(* IEC 61131-3 sources: daoli-st-library/DL_Algo (part 13) *)

(* ---- FB_DL_FirFilter.st ---- *)
(*==============================================================================
 * 组件名称 (Component)  : FB_DL_FirFilter
 * 所属子库 (Sublibrary) : DL_Algo
 * 当前版本 (Version)    : 1.0.0
 * 兼容性   (Platform)   : CODESYS 3.5+ / TwinCAT 3 / 汇川 InoProShop / 施耐德 Machine Expert
 *                         仅依赖 Standard.library（ABS），零厂商私有库
 * 功能描述 (Function)   : N 阶 FIR 直接型滤波器：抽头系数 aCoeffs[0..nTaps−1]
 *                         （aCoeffs[0] 对应最新样本，倒序卷积）：
 *                           fFiltered = Σ aCoeffs[k] × aHist[k]，k ∈ [0, nTaps−1]
 *                         样本入栈做循环移位（自深至浅倒序拷贝，防越界覆盖）。
 *                         系数和归一校验：|ΣaCoeffs − 1| < 1E-6，破约 → 锁存
 *                         故障 eCoeffSum（直流增益 ≠ 1 会引入稳态偏差，锁存
 *                         冻结输出）；N 阶钳位 [1,16]，越界钳位并置信息码
 *                         eTapsClamp；非有限样本跳过入栈并置信息码 eSampleSkip。
 * 接口     (Interface)  : 输入 fSample 输入样本、aCoeffs 抽头系数表（定长
 *                         0..15）、nTaps 有效抽头数（钳位 1~16）、bReset 复位；
 *                         输出 fFiltered 滤波输出、fCoeffSum 实测系数和
 *                         （诊断透读）、eErrCode 错误码、bError 故障标志。
 * 边界     (Boundary)   : ① **属主边界（写死）：本件只做 FIR 直接型卷积，不做
 *                         系数设计、不做 IIR 递推**；系数设计离线完成。
 *                         ② 移位：FOR 自深至浅倒序拷贝 aHist[i] := aHist[i−1]
 *                         （i ∈ [1, nTaps−1]，界宽 = 钳位后 nTaps，无越界），
 *                         aHist[0] := fSample 唯一写入点。
 *                         ③ 卷积求和界宽 = 钳位后 nTaps；aHist 尾部旧样本
 *                         （从未填充）为初值 0，首窗输出为尾零卷积（头注释
 *                         声明：上电启动期输出按零历史卷积，非异常）。
 *                         ④ 系数和归一校验在每次 nTaps 钳位后按活动抽头重算；
 *                         破约锁存后冻结输出 0（安全侧），解除沿 = bReset
 *                         上升沿（故障级码配对 bError，R45）。
 *                         ⑤ 非有限判据（R79 双判）：样本跳过（不入栈不卷积），
 *                         系数域闸含逐系数非有限判（系数 NaN 直接判归一破约
 *                         路径覆盖，另设显式非有限分支置 eCoeffSum）。
 *                         ⑥ 零全局耦合（无 GVL / VAR_EXTERNAL / 物理地址）。
 * 分工声明 (Scope)      : 与 `FB_DL_MovingAverage` 分工：等权滑动平均（FIR 特例）
 *                         归那件、任意系数 FIR 归本件；与 `FB_DL_LowPassFilter`
 *                         分工：IIR 单极点归那件。
 * 来源标签 (Source Tag) : 自研线（FIR 直接型为公开 DSP 结构 clean-room）
 * 码表     (Codes)      : 本件不占用任何全局数字码位。出口为 LREAL 组 +
 *                         ENUM 错误码；数字码位待主控收口阶段统一派号。
 * 红线自检 (Redline)    : R1 ✓ 零 GVL/VAR_EXTERNAL ｜ R2 ✓ 零 %I/%Q/%M ｜ R3 ✓ 纯 IEC 61131-3
 *                         R4 ✓ 移位界宽钳位 + 归一校验锁存 + 非有限跳过 ｜ R5 ✓ 声明逐行同行双语注释
 *                         R6 N/A（无 ENUM 状态机） ｜ R7 ✓ 一 R_TRIG 段 0 无条件刷新
 * 修订历史 (Revision)   : 2026-11-20  v1.0.0  R50 首版（批次 2 · 序号 9）
 * 验收向量 (Acceptance) : ① nTaps=2，aCoeffs=[0.5, 0.5]（Σ=1.0 过闸）：样本
 *                         序列 10, 20 → 首拍输出 0.5×10+0.5×0 = 5.0（零历史），
 *                         次拍 0.5×20+0.5×10 = 15.0，eOk；② nTaps=20 → 钳位
 *                         16，eTapsClamp；③ aCoeffs=[0.6, 0.5]（Σ=1.1）→
 *                         |1.1−1|=0.1 ≥ 1E-6 → 锁存 eCoeffSum，输出 0；
 *                         ④ 样本 NaN → uSkip 不入栈，eSampleSkip，输出不变。
 *==============================================================================*)

(*-----------------------------------------------------------------------------
 * 枚举: E_DL_FirErr（错误码；信息级不置 bError，故障级恒伴 bError=TRUE）
 *----------------------------------------------------------------------------*)
TYPE E_DL_FirErr :
(
    eOk          := 0,   // 正常 / Normal
    eCoeffSum    := 1,   // 故障级：系数和归一破约（|Σ−1| ≥ 1E-6 或含非有限） / Fault: coefficient sum not unity
    eTapsClamp   := 2,   // 信息级：抽头数越界已钳位 [1,16] / Info: tap count clamped
    eSampleSkip  := 3    // 信息级：样本非有限已跳过 / Info: non-finite sample skipped
);
END_TYPE

FUNCTION_BLOCK FB_DL_FirFilter
VAR_INPUT
    fSample : LREAL := 0.0;                    // 输入样本 [工程单位] / Input sample
    aCoeffs : ARRAY[0..15] OF LREAL;           // 抽头系数表（[0] 对应最新样本） [-] / Tap coefficients, newest-first
    nTaps   : UDINT := 4;                      // 有效抽头数，域 [1,16]（越界钳位） [个] / Active tap count
    bReset  : BOOL := FALSE;                   // 复位，上升沿清组态锁存与历史栈 [-] / Reset, rising edge clears latch and history
END_VAR
VAR_OUTPUT
    fFiltered  : LREAL;                        // 滤波输出 [工程单位] / Filtered output
    fCoeffSum  : LREAL;                        // 实测活动抽头系数和（诊断透读） [-] / Measured coefficient sum
    eErrCode   : E_DL_FirErr;                  // 错误码出口 / Error code outlet
    bError     : BOOL;                         // 故障标志（归一破约锁存） [-] / Error flag, latched
END_VAR
VAR
    _aHist    : ARRAY[0..15] OF LREAL;         // 历史样本栈（aHist[0] 最新，初值零历史） / History stack, newest first
    _nTaps    : DINT;                          // 钳位后抽头数 [个] / Clamped tap count
    _fSum     : LREAL;                         // 系数和累计中间量 [-] / Coefficient sum intermediate
    _fAcc     : LREAL;                         // 卷积累计中间量 [工程单位] / Convolution accumulator
    _bClamp   : BOOL;                          // 本拍发生抽头钳位 [-] / Tap clamp this scan
    _bNonFin  : BOOL;                          // 样本非有限当拍量 [-] / Sample non-finite this scan
    _bCoefBad : BOOL;                          // 系数归一破约当拍量 [-] / Coefficient sum violation this scan
    _bErrLatch: BOOL;                          // 归一破约锁存位（解除沿 = bReset 上升沿） / Latched coeff-sum fault
    i         : DINT;                          // 移位/卷积循环索引 / Shift and convolution loop index
    rtReset   : R_TRIG;                        // 复位沿实例，段 0 无条件调用 / Reset edge instance
END_VAR
VAR CONSTANT
    DL_FIR_NMAX   : DINT  := 16;               // 抽头定长上限 [个] / Tap count ceiling
    DL_FIR_NMIN   : DINT  := 1;                // 抽头数下限 [个] / Tap count floor
    DL_FIR_SUMTOL : LREAL := 1.0E-6;           // 系数和归一容差 [-] / Coefficient sum tolerance
    DL_FIR_ONE    : LREAL := 1.0;              // 归一目标值 [-] / Unity target
    DL_FIR_ZERO   : LREAL := 0.0;              // 判零与安全侧基准 / Zero base and safe value
END_VAR

(* —— 段 0：抽头钳位 + 非有限判 + 沿刷新 —— *)
_bClamp := FALSE;                              // 钳位量预清 / Clamp preset
_nTaps := UDINT_TO_DINT(nTaps);                // 抽头数转 DINT（越界由下步钳位） / Convert tap count
IF _nTaps > DL_FIR_NMAX THEN
    _nTaps := DL_FIR_NMAX;                     // 上越界钳 16 / Clamp high
    _bClamp := TRUE;                           // 记钳位 / Mark clamp
END_IF
IF _nTaps < DL_FIR_NMIN THEN
    _nTaps := DL_FIR_NMIN;                     // 下越界钳 1 / Clamp low
    _bClamp := TRUE;                           // 记钳位 / Mark clamp
END_IF
_bNonFin := (fSample <> fSample) OR ((fSample - fSample) <> DL_FIR_ZERO);   // 样本非有限（R79 双判） / Sample non-finite
rtReset(CLK := bReset);                        // 复位沿，每拍必调 / Reset edge, every scan

(* —— 段 1：复位沿（清锁存与历史栈） —— *)
IF rtReset.Q THEN
    _bErrLatch := FALSE;                       // 清归一破约锁存（R188 声明：解除沿 = bReset 上升沿） / Clear latch
    FOR i := 0 TO (DL_FIR_NMAX - 1) DO
        _aHist[i] := DL_FIR_ZERO;              // 清历史栈（零历史重启） / Clear history stack
    END_FOR
END_IF

(* —— 段 2：系数和归一校验（按钳位后活动抽头重算；含系数非有限判） —— *)
_fSum := DL_FIR_ZERO;                          // 系数和起步 0 / Sum start zero
FOR i := 0 TO (_nTaps - 1) DO
    _fSum := _fSum + aCoeffs[i];               // 活动抽头逐项累计 / Sum active taps
END_FOR
fCoeffSum := _fSum;                            // 透读出口 / Readout outlet
IF (_fSum <> _fSum) OR ((_fSum - _fSum) <> DL_FIR_ZERO)
   OR (ABS(_fSum - DL_FIR_ONE) >= DL_FIR_SUMTOL) THEN
    _bCoefBad := TRUE;                         // 归一破约（含系数 NaN 令和失效） / Sum violation
ELSE
    _bCoefBad := FALSE;                        // 过闸 / Pass
END_IF
IF _bCoefBad AND (NOT _bErrLatch) THEN
    _bErrLatch := TRUE;                        // 锁存（R188） / Latch
END_IF

(* —— 段 3：样本入栈（循环移位倒序拷贝，防越界；故障期/非有限期不入栈） —— *)
IF (NOT _bErrLatch) AND (NOT _bNonFin) THEN
    FOR i := (_nTaps - 1) TO DL_FIR_NMIN BY -1 DO
        _aHist[i] := _aHist[i - 1];            // 倒序拷贝（自深至浅，界宽=nTaps） / Shift down, newest-first
    END_FOR
    _aHist[0] := fSample;                      // 最新样本入栈（唯一写入点） / Push newest sample
END_IF

(* —— 段 4：卷积输出（故障安全侧 0；正常域按活动抽头求和） —— *)
IF _bErrLatch THEN
    fFiltered := DL_FIR_ZERO;                  // 归一破约冻结输出 0（安全侧，头注释④） / Frozen zero output
ELSE
    _fAcc := DL_FIR_ZERO;                      // 卷积累计起步 0 / Accumulator start
    FOR i := 0 TO (_nTaps - 1) DO
        _fAcc := _fAcc + aCoeffs[i] * _aHist[i];   // 倒序卷积逐项 / Tap-wise convolution
    END_FOR
    fFiltered := _fAcc;                        // 滤波输出 / Filtered outlet
END_IF

(* —— 段 5：出口单点映射（错误码归约，R191） —— *)
IF _bErrLatch THEN
    bError := TRUE;                            // 故障标志（R45 配对） / Error flag
    eErrCode := E_DL_FirErr.eCoeffSum;         // 故障级码 / Fault code
ELSE
    bError := FALSE;                           // 无故障级条件 / No fault
    IF _bNonFin THEN
        eErrCode := E_DL_FirErr.eSampleSkip;   // 信息级：样本跳过 / Info: skipped
    ELSIF _bClamp THEN
        eErrCode := E_DL_FirErr.eTapsClamp;    // 信息级：抽头钳位 / Info: clamped
    ELSE
        eErrCode := E_DL_FirErr.eOk;           // 正常 / Normal
    END_IF
END_IF

END_FUNCTION_BLOCK

(* ---- FB_DL_FirstOrderIdent.st ---- *)
(*
  Name        : FB_DL_FirstOrderIdent
  Category    : DL_Algo
  Version     : 1.0.0
  Purpose     : 一阶加纯滞后（FOPDT）阶跃响应回归：阶跃前后双特征点三点法估增益/时间常数/纯滞后，供自整定与 Smith 补偿取参；/ FOPDT step-response regression: two feature points before and after the step estimate gain, time constant and dead time for auto-tuning and Smith predictor
  溯源        : 自研（与 PRBS/继电器整定/扫频激励源配套），clean-room 实现
  Boundary    : ① 阶跃幅值/采样周期/窗长三重域闸，任一越域锁存故障；
                ② 辨识窗须含阶跃前稳态（>= 8 有效拍均值）与阶跃后 28.3%/63.2% 两特征点，缺任一 → 有效性 FALSE 不出参数（信息级）；
                ③ 三点法公式全代数无迭代（增益分母 = 阶跃幅值，已过正域闸；除子常量均非零）；
                ④ 非有限测量该拍不入辨识窗（窗计数暂停非快进，防污染统计）；
                ⑤ 输出 K/T/θ 非负域钳位，θ 上限 = 辨识窗时长（防无滞后误设大滞后）；
                ⑥ 本件为辨识观测层，不输出任何控制量（属主边界）。
*)
TYPE E_DL_FoiState :
(
    eIdle  := 0,                             (* 未辨识 / Not identifying *)
    eWait  := 10,                            (* 阶跃前稳态采集 / Pre-step steady sampling *)
    ePost  := 20,                            (* 阶跃后窗采集 / Post-step window sampling *)
    eReady := 30,                            (* 辨识完成（有效性查 bValid） / Finished, see bValid *)
    eFault := 90                             (* 故障锁存相 / Fault latched *)
);
END_TYPE

TYPE E_DL_FoiCause :
(
    eNone      := 0,                         (* 无成因 / No cause *)
    eCfgIllegal:= 1,                        (* 组态非法：幅值/周期/窗长越域 / Illegal config *)
    eNoFeat    := 2,                        (* 信息级：缺稳态/特征点或增益反号 / Info: feature missing *)
    ePhaseBad  := 3                         (* 非法相位兜底 / Illegal phase fallback *)
);
END_TYPE

FUNCTION_BLOCK FB_DL_FirstOrderIdent
VAR_INPUT
    fMeas   : REAL := 0.0;                   (* 回路测量值（任意工程量）[-] / Loop measurement *)
    fStepAmp: REAL := 10.0;                  (* 阶跃幅值，域 > 0 [工程单位] / Step amplitude *)
    tSample : TIME := T#100MS;               (* 采样周期，域 > T#0S [ms] / Sampling period *)
    nWin    : INT := 128;                    (* 阶跃后窗长，域 20..256 [拍] / Post-step window length *)
    bStart  : BOOL := FALSE;                 (* 启动辨识命令，上升沿进入稳态采集 [-] / Start command *)
    bEnable : BOOL := TRUE;                  (* 使能 [-] / Enable *)
    bReset  : BOOL := FALSE;                 (* 复位命令，上升沿清故障与结果 [-] / Reset command *)
END_VAR
VAR_OUTPUT
    fK      : REAL;                          (* 增益出口 = 稳态增量 / 阶跃幅值 [-] / Gain outlet *)
    fTau    : REAL;                          (* 时间常数出口 [s] / Time constant outlet *)
    fTheta  : REAL;                          (* 纯滞后出口（非负，上限 = 窗时长）[s] / Dead time outlet *)
    bValid  : BOOL;                          (* 结果有效性出口 [-] / Result validity *)
    nSamples: INT;                           (* 阶跃后窗内有效样本数 [拍] / Valid samples in window *)
    eState  : E_DL_FoiState;                 (* 状态出口 / State outlet *)
    eCause  : E_DL_FoiCause;                 (* 成因出口（R190 归因唯一） / Cause outlet *)
    bError  : BOOL;                          (* 故障锁存标志 [-] / Fault latch flag *)
END_VAR
VAR
    _eState : E_DL_FoiState := E_DL_FoiState.eIdle;  (* 内部相位（CASE 唯一写入目标） / Internal phase *)
    _eCause : E_DL_FoiCause := E_DL_FoiCause.eNone;  (* 成因锁存量 / Latched cause *)
    rtStart : R_TRIG;                        (* 启动沿实例，段 0 无条件调用 / Start edge instance *)
    rtReset : R_TRIG;                        (* 复位沿实例，段 0 无条件调用 / Reset edge instance *)
    _bFault : BOOL;                          (* 故障锁存位 / Latched fault bit *)
    _bCfgBad: BOOL;                          (* 组态非法当拍量 / Illegal config this scan *)
    _bFin   : BOOL;                          (* 测量有限性当拍量（边界④） / Measurement finiteness *)
    _nWinE  : INT;                           (* 钳位后生效窗长 [拍] / Effective window length *)
    _nPreN  : INT;                           (* 稳态已采有效拍数 [拍] / Pre samples collected *)
    _fPreSum: REAL;                          (* 稳态样本累加和 [工程单位] / Pre samples sum *)
    _fY0    : REAL;                          (* 阶跃前稳态均值 [工程单位] / Baseline mean *)
    _nRecN  : INT;                           (* 窗内已收有效样本数 [拍] / Window samples count *)
    _aRec   : ARRAY[1..256] OF REAL;         (* 窗内样本记录（连续有效区）[工程单位] / Window sample record *)
    _fYinf  : REAL;                          (* 窗末稳态均值 [工程单位] / Final steady mean *)
    _fDelta : REAL;                          (* 稳态增量中间量 [工程单位] / Steady delta *)
    _fKI    : REAL;                          (* 增益中间量 [-] / Gain intermediate *)
    _fT1    : REAL;                          (* 28.3% 特征时刻 [s] / Feature time 1 *)
    _fT2    : REAL;                          (* 63.2% 特征时刻 [s] / Feature time 2 *)
    _fTauI  : REAL;                          (* 时间常数中间量 [s] / Tau intermediate *)
    _fThI   : REAL;                          (* 滞后中间量 [s] / Theta intermediate *)
    _i      : INT;                           (* 窗扫描游标 [拍] / Window scan cursor *)
    _fDtSec : REAL;                          (* 采样周期秒值，域 > eps [s] / Sampling period seconds *)
END_VAR
VAR CONSTANT
    DL_FOI_NPRE   : INT  := 8;               (* 阶跃前稳态最少有效拍数（边界②）[拍] / Pre-step minimum samples *)
    DL_FOI_NTAIL  : INT  := 8;               (* 窗末稳态平均样本数 [拍] / Tail averaging samples *)
    DL_FOI_WMIN   : INT  := 20;              (* 窗长下限（边界①）[拍] / Window lower bound *)
    DL_FOI_WMAX   : INT  := 256;             (* 窗长上限（数组容量）[拍] / Window upper bound *)
    DL_FOI_EPS    : REAL := 1.0E-6;          (* 判零容差 [-] / Epsilon *)
    DL_FOI_L1     : REAL := 0.283;           (* 特征点 1 归一化水平（1-exp(-1/3)）[-] / Feature level 1 *)
    DL_FOI_L2     : REAL := 0.632;           (* 特征点 2 归一化水平（1-exp(-1)）[-] / Feature level 2 *)
    DL_FOI_STEPDET: REAL := 0.1;             (* 阶跃检测阈（幅值占比）[-] / Step detect threshold *)
END_VAR

(* —— 段 0：当拍判据派生 + 实例无条件刷新（R228A） —— *)
_fDtSec := TIME_TO_LREAL(tSample) / 1000.0;              (* 采样周期秒化（除子常量 1000） / Sampling period seconds *)
_bCfgBad := (fStepAmp <= DL_FOI_EPS)                     (* 阶跃幅值正域闸（边界①） / Step amplitude gate *)
            OR NOT (tSample > T#0S)                      (* 采样周期正域闸（边界①） / Sampling gate *)
            OR (nWin < DL_FOI_WMIN) OR (nWin > DL_FOI_WMAX);   (* 窗长域闸（边界①） / Window gate *)
rtStart(CLK := bStart);                                  (* 启动沿每拍必调 / Start edge every scan *)
rtReset(CLK := bReset);                                  (* 复位沿每拍必调 / Reset edge every scan *)
_bFin := (fMeas = fMeas) AND ((fMeas - fMeas) = (fMeas - fMeas));   (* 测量 NaN 自反 + Inf 差判闸（边界④） / Measurement NaN and Inf gate *)
_nWinE := nWin;                                          (* 生效窗长初值 / Effective window init *)
IF _nWinE < DL_FOI_WMIN THEN
    _nWinE := DL_FOI_WMIN;                               (* 窗长下限钳位 / Window lower clamp *)
END_IF
IF _nWinE > DL_FOI_WMAX THEN
    _nWinE := DL_FOI_WMAX;                               (* 窗长上限钳位（防数组越界） / Window upper clamp *)
END_IF

(* —— 段 1：单拍量预清零（R107） —— *)
nSamples := 0;                                           (* 样本数出口预清（派生拍覆盖） / Samples outlet preset *)

(* —— 段 2：复位沿处理（作用域：清故障 + 清辨识状态 + 迁 eIdle，R283 逐项声明） —— *)
IF rtReset.Q THEN
    _bFault := FALSE;                                    (* 清故障锁存 / Clear fault *)
    _eCause := E_DL_FoiCause.eNone;                      (* 清成因 / Clear cause *)
    bValid := FALSE;                                     (* 清有效性出口 / Clear validity *)
    fK := 0.0; fTau := 0.0; fTheta := 0.0;               (* 清 K/T/θ 出口 / Clear K T theta *)
    _nPreN := 0; _fPreSum := 0.0;                        (* 清稳态采集量 / Clear pre sampling *)
    _nRecN := 0;                                         (* 清窗样本数 / Clear window count *)
    _eState := E_DL_FoiState.eIdle;                      (* 迁未辨识相 / Back to idle *)
END_IF

(* —— 段 3：组态故障锁存（锁存至复位沿，R189） —— *)
IF _bCfgBad AND NOT _bFault THEN
    _bFault := TRUE;                                     (* 锁存故障位 / Latch fault *)
    _eCause := E_DL_FoiCause.eCfgIllegal;                (* 成因：组态非法 / Cause illegal config *)
    _eState := E_DL_FoiState.eFault;                     (* 同步迁故障相 / Migrate to fault *)
END_IF

(* —— 段 4：CASE 主状态机（ELSE 兜底迁 eFault，红线 6） —— *)
CASE _eState OF
    E_DL_FoiState.eIdle:                                 (* 未辨识：出口保持确定值 / Idle *)
        bValid := FALSE;                                 (* 未辨识有效性 FALSE（不留陈旧） / Validity false *)
        IF rtStart.Q AND bEnable AND NOT _bFault THEN
            _nPreN := 0; _fPreSum := 0.0;                (* 清稳态采集（新一轮） / Clear pre sampling *)
            _nRecN := 0;                                 (* 清窗样本（新一轮） / Clear window samples *)
            _eState := E_DL_FoiState.eWait;              (* 进入稳态采集相 / Enter pre sampling *)
        END_IF
    E_DL_FoiState.eWait:                                 (* 稳态采集相：阶跃前基线 / Pre-step sampling *)
        IF NOT bEnable THEN
            _eState := E_DL_FoiState.eIdle;              (* 失能回未辨识 / Back to idle *)
        ELSIF _bFin THEN                                 (* 非有限拍不入窗（计数暂停，边界④） / Skip non-finite *)
            _fPreSum := _fPreSum + fMeas;                (* 稳态样本累加 / Pre sample accumulate *)
            _nPreN := _nPreN + 1;                        (* 有效拍数净额 +1 / Valid count *)
            IF _nPreN >= DL_FOI_NPRE THEN
                _fY0 := _fPreSum / INT_TO_REAL(_nPreN);  (* 稳态均值（除子 = 有效拍数 >= 8） / Baseline mean *)
                IF ABS(fMeas - _fY0) > DL_FOI_STEPDET * fStepAmp THEN   (* 阶跃检测（幅值占比直比） / Step detected *)
                    _nRecN := 0;                         (* 窗样本从阶跃后重计 / Window from step *)
                    _eState := E_DL_FoiState.ePost;      (* 进入阶跃后窗相 / Enter post window *)
                END_IF
            END_IF
        END_IF
    E_DL_FoiState.ePost:                                 (* 阶跃后窗相：连续采样至窗满 / Post window *)
        IF NOT bEnable THEN
            _eState := E_DL_FoiState.eIdle;              (* 失能回未辨识 / Back to idle *)
        ELSIF _bFin THEN                                 (* 非有限拍不入窗（暂停非快进，边界④） / Skip non-finite *)
            IF _nRecN < _nWinE THEN
                _nRecN := _nRecN + 1;                    (* 窗样本净额 +1（写入点下标域内） / Window count *)
                _aRec[_nRecN] := fMeas;                  (* 样本入记录（下标 1.._nWinE 钳定） / Sample recorded *)
            END_IF
            IF _nRecN >= _nWinE THEN
                nSamples := _nRecN;                      (* 窗内有效样本数出口 / Samples outlet *)
                _fYinf := 0.0;                           (* 窗末均值累加清零 / Tail mean clear *)
                FOR _i := _nRecN - DL_FOI_NTAIL + 1 TO _nRecN DO   (* 末 8 样本均值（区段域内） / Tail mean *)
                    _fYinf := _fYinf + _aRec[_i];        (* 尾段累加 / Tail accumulate *)
                END_FOR
                _fYinf := _fYinf / INT_TO_REAL(DL_FOI_NTAIL);   (* 尾段均值（除子常量 8） / Tail mean *)
                _fDelta := _fYinf - _fY0;                (* 稳态增量（阶跃后末均值 - 阶跃前均值） / Steady delta *)
                _fKI := _fDelta / fStepAmp;              (* 增益（除子 = 幅值已过正域闸，边界③） / Gain *)
                _fT1 := 0.0; _fT2 := 0.0;                (* 特征时刻清零（未命中哨兵） / Feature times clear *)
                FOR _i := 1 TO _nRecN DO
                    IF (_fT1 <= DL_FOI_EPS) AND (_aRec[_i] >= _fY0 + DL_FOI_L1 * _fDelta) THEN
                        _fT1 := INT_TO_REAL(_i) * _fDtSec;   (* 首过 28.3% 时刻（边界②） / First level 1 time *)
                    END_IF
                    IF (_fT2 <= DL_FOI_EPS) AND (_aRec[_i] >= _fY0 + DL_FOI_L2 * _fDelta) THEN
                        _fT2 := INT_TO_REAL(_i) * _fDtSec;   (* 首过 63.2% 时刻（边界②） / First level 2 time *)
                    END_IF
                END_FOR
                IF (_fT1 > DL_FOI_EPS) AND (_fT2 > DL_FOI_EPS) AND (_fT2 > _fT1) AND (_fKI > 0.0) THEN
                    _fTauI := 1.5 * (_fT2 - _fT1);       (* 两点法时间常数（公开代数式，除子常量） / Two-point tau *)
                    _fThI := _fT2 - _fTauI;              (* 两点法纯滞后 / Two-point theta *)
                    IF _fTauI < 0.0 THEN
                        _fTauI := 0.0;                   (* 时间常数非负钳位（边界⑤） / Tau clamp *)
                    END_IF
                    IF _fThI < 0.0 THEN
                        _fThI := 0.0;                    (* 滞后非负钳位（边界⑤） / Theta clamp *)
                    END_IF
                    IF _fThI > INT_TO_REAL(_nRecN) * _fDtSec THEN
                        _fThI := INT_TO_REAL(_nRecN) * _fDtSec;   (* 滞后上限 = 窗时长（边界⑤） / Theta window cap *)
                    END_IF
                    fK := _fKI;                          (* 增益出口（非负已闸） / Gain outlet *)
                    fTau := _fTauI;                      (* 时间常数出口 / Tau outlet *)
                    fTheta := _fThI;                     (* 滞后出口 / Theta outlet *)
                    bValid := TRUE;                      (* 有效性 TRUE / Validity true *)
                    _eState := E_DL_FoiState.eReady;     (* 迁完成相 / To ready *)
                ELSE
                    bValid := FALSE;                     (* 缺特征点或增益反号：不出参数（边界②⑤） / Invalid *)
                    _eCause := E_DL_FoiCause.eNoFeat;    (* 信息级成因（不置 bError） / Info cause *)
                    _eState := E_DL_FoiState.eReady;     (* 迁完成相（无效结论） / To ready invalid *)
                END_IF
            END_IF
        END_IF
    E_DL_FoiState.eReady:                                (* 完成相：结论冻结保持 / Ready *)
        IF rtStart.Q THEN
            _eState := E_DL_FoiState.eIdle;              (* 新启动沿经 eIdle 重入（防隐性回夹） / Restart via idle *)
        END_IF
    E_DL_FoiState.eFault:                                (* 故障相：冻结保持，仅复位沿出 / Fault *)
        ;                                                (* 锁存回放（R28） / Replay from latch *)
    ELSE                                                 (* 非法相位兜底迁安全态 / Illegal phase fallback *)
        _eState := E_DL_FoiState.eFault; _bFault := TRUE;    (* 迁故障相 + 同步锁存 / To fault and latch *)
        _eCause := E_DL_FoiCause.ePhaseBad;              (* 成因：非法相位 / Cause illegal phase *)
END_CASE

(* —— 段 5：出口映射（bError/eState 同源，R191） —— *)
bError := _bFault;                                       (* 故障标志镜像 / Fault flag mirror *)
eState := _eState;                                       (* 状态出口 / State outlet *)
eCause := _eCause;                                       (* 成因出口 / Cause outlet *)
END_FUNCTION_BLOCK

(* ---- FB_DL_FlowSqrtExtract.st ---- *)
(*
    FB_DL_FlowSqrtExtract —— 差压流量开方 + 小信号切除
    ------------------------------------------------------------------
    分类      : DL_Algo / ProcessControl
    前缀      : FB_DL_
    版本      : 1.0.0
    溯源      : 差压式流量测量的公开仪表工程惯例（开方 + 小信号切除 + 一阶阻尼 + 满量程标定）；
                只借「阻尼与限幅同层」的组织方式，迟滞切除判据、阻尼律、错误分级、
                状态组织与码位 100% 自有；开方一律委托平台内建 SQRT，禁牛顿迭代重实现；
                clean-room 重写，未复制任何闭源厂商源码，参考实现仅限 MIT/Apache 许可
    平台      : 纯 IEC 61131-3，CODESYS V3.5+ / TwinCAT 3 / InoProShop 通用
    作者      : 道莅代码库 · PLC编程专家（R19）
    ------------------------------------------------------------------
    功能说明  : 孔板流量在 5% 以下差压时开方后噪声被放大 4~5 倍，HMI 上流量在零附近乱跳，
                操作工据此判「有没有流量」必然误判；硬切又在切点附近反复跳。
                本件把「迟滞切除」做进块内：进入切除要跌破「切除点 − 迟滞带宽」，
                退出切除要重新越过切除点，带内保持上一状态（本件核心防御，与硬切的分界）。
                其余防御：① 量程与采样周期非法即故障级 2710，输出 0；
                ② 差压负漂取 0 参与运算（直接开方会出 NaN）并置信息码；
                ③ 差压非有限即故障级 2711，保持末次有效输出——零流量与信号故障
                   在联锁上是两个结论，绝不输出 0；
                ④ 输出双侧钳位（下 0，上 fFlowSpan），超顶置 bSaturated。
                职责边界：本件只出流量工程量，不做温压补偿（归补偿件），不做累积。
    错误码    : 16#0002_2701 切除点超域已钳位 / 差压负漂已取 0 / 切除迟滞带保持中——信息级，正常防御
                16#0002_2702 预留禁用（信息级，不得挪用）
                16#0002_2710 量程或采样周期参数非法——故障级，输出 0 且 bValid = FALSE
                16#0002_2711 差压输入非有限——故障级，保持末次有效输出且 bValid = FALSE
                16#0002_2712 预留禁用（故障级，不得挪用）
    码位总账  : 16#0002_2701 用 / 16#0002_2702 预留 ｜ 16#0002_2710 用 / 16#0002_2711 用 / 16#0002_2712 预留
    状态机    : R6 标注 N/A —— 本组件为纯函数无顺序状态机，无 CASE 可写，非法状态不可能出现
                （切除态由单比特锁存 bCutLatch 承载，非顺序状态机）
    采样约定  : fbTrigReset 在本体首部无条件刷新；阻尼系数 α 隐含以 tSampleTime 为步长，
                采样周期未知或越域时阻尼律不可信，故并入 2710 判据（tSampleTime 越域即故障）。
    修订记录  : 2026-11-16 v1.0.0 首次入库（R19）
*)
FUNCTION_BLOCK FB_DL_FlowSqrtExtract
VAR_INPUT
    bEnable        : BOOL;                    // 使能，FALSE 输出 0 并冻结阻尼状态 / enable, FALSE outputs zero and freezes the damping state
    bReset         : BOOL;                    // 复位，上升沿清阻尼状态与切除锁存 / reset, rising edge clears the damping state and the cutoff latch
    fDp            : REAL := 0.0;             // 差压输入 [用户单位]，范围 -10.0~110.0 / differential pressure input [user unit], range -10.0~110.0
    fDpSpan        : REAL := 100.0;           // 差压满量程 [用户单位]，必须 > 0 / differential pressure span [user unit], must be > 0
    fFlowSpan      : REAL := 100.0;           // 流量满量程 [m3/h]，必须 > 0 / flow span [m3/h], must be > 0
    fCutPercent    : REAL := 1.0;             // 切除点（差压满量程百分比）[%]，范围 0.0~20.0，0 = 不切除 / cutoff point as a percentage of the span [%], range 0.0~20.0, zero disables it
    fCutHystPercent : REAL := 0.3;            // 切除迟滞带宽度（相对满量程）[%]，范围 0.0~10.0 / hysteresis band width of the cutoff relative to the span [%], range 0.0~10.0
    fDampCoef      : REAL := 0.2;             // 一阶阻尼系数 α [无量纲]，范围 0.0~1.0，0 = 不阻尼，1 = 冻结 / first order damping factor [dimensionless], 0.0~1.0
    tSampleTime    : TIME := T#100MS;         // 采样周期 [ms]，范围 1~10000 / sample time [ms], range 1~10000
    bSquareRoot    : BOOL := TRUE;            // TRUE = 开方（差压型），FALSE = 线性（已开方变送器）/ TRUE takes the square root, FALSE is linear
END_VAR
VAR_OUTPUT
    fFlow          : REAL;                    // 输出流量 [m3/h]，范围 0.0~fFlowSpan / output flow [m3/h], range 0.0~fFlowSpan
    bCutoff        : BOOL;                    // 当前处于切除区，输出被强制 0 / currently inside the cutoff band, output forced to zero
    bSaturated     : BOOL;                    // 输出被满量程钳位 / output clamped at the span
    uCutCount      : UDINT;                   // 切除进入次数，抖动监视用 [次] / cutoff entries for chatter monitoring [times]
    eErr           : UDINT;                   // 错误码，0=正常 / error id, 0=ok
    bError         : BOOL;                    // 故障标志，eErr 为故障级时 TRUE / error flag, TRUE on fault-level eErr
    bValid         : BOOL;                    // 输出是否可用 / output valid flag
END_VAR
VAR
    fbTrigReset    : R_TRIG;                  // 复位上升沿实例，本体首部无条件刷新 / reset edge instance, refreshed unconditionally
    bCutLatch      : BOOL;                    // 切除锁存（带内保持上一状态）/ cutoff latch, holds the previous state inside the band
    fDamped        : REAL;                    // 一阶阻尼内部状态 [m3/h] / first order damping internal state [m3/h]
    fRatio         : REAL;                    // 差压/满量程归一比值 [无量纲]，范围 0.0~1.0 / normalised ratio [dimensionless], range 0.0~1.0
    fRaw            : REAL;                   // 切除与阻尼前的瞬时流量 [m3/h] / instantaneous flow before cutoff and damping [m3/h]
    fDpEff         : REAL;                    // 负漂修正后的差压 [用户单位] / differential pressure after the negative drift correction [user unit]
    fCutEff        : REAL;                    // 域钳位后的切除点 [%] / cutoff point after domain clamping [%]
    fHystEff       : REAL;                    // 域钳位后的迟滞带宽度 [%] / hysteresis band width after domain clamping [%]
    fDampEff       : REAL;                    // 域钳位后的阻尼系数 [无量纲] / damping factor after domain clamping [dimensionless]
    bNonFin        : BOOL;                    // 输入非有限判定标志 / non-finite input flag
    bEnterCut      : BOOL;                    // 本拍新进入切除区（用于计数）/ newly entered the cutoff band in this cycle, used for counting
END_VAR
VAR CONSTANT
    DL_FSQ_CUT_MAX   : REAL := 20.0;          // 切除点上限 [%] / cutoff point upper bound [%]
    DL_FSQ_HYST_MAX  : REAL := 10.0;          // 迟滞带宽度上限 [%] / hysteresis band width upper bound [%]
    DL_FSQ_DAMP_MAX  : REAL := 1.0;           // 阻尼系数上限 [无量纲] / damping factor upper bound [dimensionless]
    DL_FSQ_DT_MAX    : TIME := T#10S;         // 采样周期上限 [ms] / sample time upper bound [ms]
    DL_FSQ_DT_MIN    : TIME := T#1MS;         // 采样周期下限 [ms] / sample time lower bound [ms]
    DL_FLOAT_EPS     : REAL := 1.0E-6;        // 浮点判等容差 [无量纲] / float equality tolerance [dimensionless]
    DL_FSQ_PERCENT   : REAL := 100.0;         // 百分比换算因子 [%] / percent conversion factor [%]
    DL_FSQ_RATIO_MAX : REAL := 1.0;           // 归一比值上限 [无量纲] / normalised ratio upper bound [dimensionless]
    DL_FSQ_INF_GUARD : REAL := 1.0E38;        // 非有限幅值判定阈值 [无量纲] / non-finite magnitude guard [dimensionless]
    DL_FSQ_CNT_MAX   : UDINT := 16#FFFF_FFFE; // 切除计数饱和值 [次] / cutoff counter saturation value [times]
    DL_FSQ_ZERO      : REAL := 0.0;           // 零值常量，避免裸字面量 [无量纲] / zero constant, avoids a bare literal [dimensionless]
END_VAR

// 段 1｜边沿实例无条件周期刷新（红线：严禁放入条件分支）/ segment 1, unconditional edge refresh
fbTrigReset(CLK := bReset);

// 段 2｜输出与错误状态预置（fFlow 不预置，非有限时须保持末次有效值）/ segment 2, preset outputs except the held flow
eErr := 0;                                    // 预置无错误 / preset no error
bError := FALSE;                              // 预置无故障 / preset no fault
bValid := FALSE;                              // 预置不可用 / preset invalid
bSaturated := FALSE;                          // 预置未饱和 / preset not saturated
bCutoff := FALSE;                             // 预置非切除态 / preset outside the cutoff band
bEnterCut := FALSE;                           // 预置非新进切除 / preset not entering the cutoff band

// 段 3｜使能闸：失能输出 0 并冻结阻尼状态 / segment 3, enable gate
IF NOT bEnable THEN
    fFlow := DL_FSQ_ZERO;                     // 失能输出 0 [m3/h] / output zero while disabled [m3/h]
    RETURN;                                   // 失能即出口，阻尼状态自然冻结 / disabled is the exit, the damping state stays frozen
END_IF

// 段 4｜参数闸：量程、采样周期、参数有限性（隐含阻尼律的时基前提）/ segment 4, parameter gate
bNonFin := (fDpSpan <> fDpSpan) OR (fDpSpan > DL_FSQ_INF_GUARD) OR (fDpSpan < -DL_FSQ_INF_GUARD)
        OR (fFlowSpan <> fFlowSpan) OR (fFlowSpan > DL_FSQ_INF_GUARD) OR (fFlowSpan < -DL_FSQ_INF_GUARD); // 参数非有限判定 / parameter non-finite detection
IF bNonFin OR (fDpSpan <= DL_FLOAT_EPS) OR (fFlowSpan <= DL_FLOAT_EPS)
   OR (tSampleTime < DL_FSQ_DT_MIN) OR (tSampleTime > DL_FSQ_DT_MAX) THEN
    eErr := 16#0002_2710;                     // 量程或采样周期非法故障码 / span or sample time fault id
    bError := TRUE;                           // 置故障标志 / raise the error flag
    fFlow := DL_FSQ_ZERO;                     // 参数非法时输出 0 / output zero when the parameters are illegal
    bValid := FALSE;                          // 输出不可用 / output not usable
    RETURN;                                   // 故障级提前返回 / early return on fault
END_IF

// 段 5｜差压输入非有限闸：保持末次有效输出，绝不输出 0 / segment 5, non-finite dp gate
IF (fDp <> fDp) OR (fDp > DL_FSQ_INF_GUARD) OR (fDp < -DL_FSQ_INF_GUARD) THEN
    eErr := 16#0002_2711;                     // 输入非有限故障码 / non-finite input fault id
    bError := TRUE;                           // 置故障标志 / raise the error flag
    bValid := FALSE;                          // 输出不可用 / output not usable
    RETURN;                                   // 保持末次 fFlow，零流量与信号故障是两个结论 / keep the last flow, zero flow and a signal fault are two different conclusions
END_IF

// 段 6｜参数域钳位（切除点、迟滞带、阻尼系数各自收敛）/ segment 6, parameter domain clamp
fCutEff := MIN(MAX(fCutPercent, DL_FSQ_ZERO), DL_FSQ_CUT_MAX);   // 切除点收敛到 0.0~20.0 % / converge the cutoff into 0.0~20.0 %
fHystEff := MIN(MAX(fCutHystPercent, DL_FSQ_ZERO), DL_FSQ_HYST_MAX); // 迟滞带宽收敛到 0.0~10.0 % / converge the hysteresis band into 0.0~10.0 %
fDampEff := MIN(MAX(fDampCoef, DL_FSQ_ZERO), DL_FSQ_DAMP_MAX);   // 阻尼系数收敛到 0.0~1.0 / converge the damping factor into 0.0~1.0
IF (fCutPercent > DL_FSQ_CUT_MAX) OR (fCutPercent < DL_FSQ_ZERO) THEN
    eErr := 16#0002_2701;                     // 信息级：切除点超域已钳位 / info level, the cutoff point was clamped
END_IF

// 段 7｜负漂修正：差压变送器零点负漂是常态，直接开方会出 NaN / segment 7, negative drift correction
fDpEff := fDp;                                // 取入参副本 / copy the input
IF fDpEff < DL_FSQ_ZERO THEN
    fDpEff := DL_FSQ_ZERO;                    // 负漂取 0 参与运算 / clamp a negative drift to zero before the square root
    eErr := 16#0002_2701;                     // 信息级：负漂已取 0 / info level, the negative drift was clamped
END_IF

// 段 8｜复位沿清阻尼与切除锁存（在切除判定之前生效）/ segment 8, reset clears the damping state and the latch
IF fbTrigReset.Q THEN
    fDamped := DL_FSQ_ZERO;                   // 清阻尼内部状态 / clear the damping state
    bCutLatch := FALSE;                       // 清切除锁存 / clear the cutoff latch
END_IF

// 段 9｜归一比值与瞬时流量（开方委托内建，入参已保证非负）/ segment 9, ratio and instantaneous flow
fRatio := fDpEff / fDpSpan;                   // 满量程已由段 4 保证 > 0，除法安全 / the span is positive by segment 4, the division is safe
fRatio := MIN(MAX(fRatio, DL_FSQ_ZERO), DL_FSQ_RATIO_MAX); // 比值双侧钳位到 0.0~1.0 / clamp the ratio into 0.0~1.0
IF bSquareRoot THEN
    fRaw := SQRT(fRatio) * fFlowSpan;         // 开方型：委托内建 SQRT [m3/h] / square root type, delegate to the built-in SQRT [m3/h]
ELSE
    fRaw := fRatio * fFlowSpan;               // 线性型：已开方变送器只做切除与阻尼 [m3/h] / linear type, only cutoff and damping [m3/h]
END_IF

// 段 10｜迟滞切除（核心防御）：退出要越过切除点，进入要跌破切除点减带宽 / segment 10, hysteresis cutoff
IF fCutEff <= DL_FLOAT_EPS THEN
    bCutLatch := FALSE;                       // 切除点 0 = 不切除 / a zero cutoff point disables the function
ELSE
    IF (fRatio * DL_FSQ_PERCENT) >= fCutEff THEN
        bCutLatch := FALSE;                   // 越过切除点即退出切除 / leaving the cutoff once the point is crossed again
    ELSIF (fRatio * DL_FSQ_PERCENT) < (fCutEff - fHystEff) THEN
        IF NOT bCutLatch THEN
            bEnterCut := TRUE;                // 新进入切除区，用于计数 / newly entered, used for counting
        END_IF
        bCutLatch := TRUE;                    // 跌破「切除点 − 带宽」才进入切除 / entering only below the point minus the band
    END_IF
END_IF
bCutoff := bCutLatch;                         // 对外发布切除态 / publish the cutoff state
IF bCutLatch THEN
    fRaw := DL_FSQ_ZERO;                      // 切除区强制 0，抑制开方噪声放大 / force zero inside the cutoff band to suppress noise amplification
END_IF

// 段 11｜切除进入计数（饱和，抖动监视）/ segment 11, saturating cutoff entry counter
IF bEnterCut AND (uCutCount < DL_FSQ_CNT_MAX) THEN
    uCutCount := uCutCount + 1;               // 饱和加一，绝不回绕 / saturating increment, never wraps
END_IF

// 段 12｜一阶阻尼（α = 1 等价冻结，α = 0 直通）/ segment 12, first order damping
fDamped := fDamped + fDampEff * (fRaw - fDamped); // 一阶离散阻尼 [m3/h] / first order discrete damping [m3/h]

// 段 13｜输出双侧钳位（只做单侧是常见缺陷）/ segment 13, two-sided output clamp
fFlow := fDamped;                             // 先取阻尼输出 / take the damped value first
IF fFlow > fFlowSpan THEN
    fFlow := fFlowSpan;                       // 上限钳位 / clamp at the upper bound
    bSaturated := TRUE;                       // 标记饱和 / flag the saturation
ELSIF fFlow < DL_FSQ_ZERO THEN
    fFlow := DL_FSQ_ZERO;                     // 下限钳位 / clamp at the lower bound
END_IF

// 段 14｜发布状态（信息码永不置 bError）/ segment 14, publish the status
bValid := TRUE;                               // 通过全部闸门，输出可用 / all gates passed, the output is usable
bError := FALSE;                              // 信息级不置故障 / info level never raises a fault
END_FUNCTION_BLOCK

(* ---- FB_DL_FopdtStepIdent.st ---- *)
(*
  ==================================================================
  组件名 Component  : FB_DL_FopdtStepIdent
  分类   Category   : DL_Algo
  版本   Version    : 1.0.1
  功能   Purpose    : 阶跃响应 FOPDT（一阶惯性 + 纯延迟）参数辨识，供 PID 整定使用。
                      阶跃窗内「时刻 + 过程量」二元组以环窗缓存，稳定或超时后按
                      时间序遍历样本，两条 clean-room 方法并行求解并在出口二选一：
                      一 两点法：取 28.3% 与 63.2% 两个穿越点，
                         T = 1.5 * (t63 - t28)，L = t63 - T；
                      二 切线法：取最大斜率点切线，
                         T = ΔPV / 最大斜率，L = t_slope - (PV_slope - PV_base) / 带符号斜率
                         （斜率符号取 SIGN(ΔPV)，负向阶跃与两点法同口径）；
                      增益 K = ΔPV / ΔMV 两法共用。
  溯源   Origin     : 阶跃辨识两点法与切线法均为公开控制工程方法；本件为 clean-room
                      实现，仅借鉴来源分类与参数域组织（来源标签 t2-5-modpid 的 PID
                      自整定概念域），未复制任何闭源代码行。
  平台   Platform   : 纯 IEC 61131-3（TON / R_TRIG / REAL 运算，无私有库、无方言转换）
  作者   Author     : 道莅代码库 · PLC 编程专家（R55）
  ------------------------------------------------------------------
  同拍双窗配比约束（R100）：tSettle 必须小于 tTimeout —— 稳定确认窗短于相超时窗，
                      两窗职责分离：tSettle 判「可以进入评估」，tTimeout 判「辨识失败退出」，
                      任一窗不得兼作另一窗用途；配比反置在组态域闸内直接判故障。
  边界 Boundary     :
                      一 本件只输出辨识参数与有效性，不算 PID 参数、不写调节器（属主边界）；
                      二 环窗遍历一律按时间序（自最旧样本起），禁按数组下标序（R194）；
                      三 采样拍周期由引脚 fSampleS 给出（秒），不读系统时基；
                      四 故障锁存解除路径 = bReset 上升沿 或 bEnable 下降沿，两条均恒可达；
                      五 无全局变量、无外部变量声明、无物理地址寻址。
  输出契约 Output contract:
                      fGainK / fTauS / fDeadS 仅在 bValid 为真拍更新，其余拍保持上一次
                      成功辨识值；非有限中间结果一律不写入出口（出口保持上拍值）；
                      bIdentDone 为单拍脉冲（内部 _bIdentInt 置位、统一出口映射后撤销，
                      R187 两段式）；eCause 各成因独立成员（R190 归因唯一）。
  修订记录 Revision  :
    2026-11-20  v1.0.0  R55 首版（批 1 · 序号 2）
    2026-11-20  v1.0.1  R56 返修（7.2）：切线法截距改用带符号斜率 _fSlopeSig（符号取
                        SIGN(_fDeltaPv)，量级守卫仍由 _fSlopeMax > DL_FOPDT_EPS 证明），
                        负向阶跃不再系统性高估死区时间；eDone 相重启分支补清
                        _fPvSlopeMax / _fTSlopeMax（与 eIdle 分支对齐）。
  ==================================================================
*)

TYPE E_DL_FopdtState :
(
    eIdle    := 0,      // 空闲：等待阶跃上升沿 / idle, waiting for the step rising edge
    eRise    := 10,     // 上升：缓存样本并监视稳定 / rising, buffering samples and watching settle
    eEval    := 20,     // 评估：时间序遍历样本算参数 / evaluating, traversing samples in time order
    eDone    := 30,     // 完成：参数已交付并驻留 / done, parameters delivered and held
    eFault   := 90      // 故障：原因锁存 / fault, cause latched
);
END_TYPE

TYPE E_DL_FopdtCause :
(
    eNone       := 0,   // 无成因 / no cause
    eCfgIllegal := 1,   // 组态非法：阈值或采样周期越域 / illegal config, threshold or sample period out of domain
    eMvZero     := 2,   // 阶跃幅度近零，增益不可算 / step amplitude near zero, gain not computable
    eLackResp   := 3,   // 响应不足：总变化未达最小可辨量 / response too small, total change below the floor
    eNoSettle   := 4,   // 超时未稳定 / timeout without settle
    eNoCross    := 5,   // 未捕获穿越点或样本不足 / crossing points missing or too few samples
    eDeadNeg    := 6,   // 纯延迟算出负值，已按零处理（信息级）/ dead time negative and forced to zero, informational
    ePhaseBad   := 7    // 非法相位兜底 / illegal phase fallback
);
END_TYPE

FUNCTION_BLOCK FB_DL_FopdtStepIdent
VAR_INPUT
    bEnable        : BOOL := TRUE;           // 使能，下降沿清状态回空闲 [-] / enable, falling edge clears the state back to idle
    bReset         : BOOL := FALSE;          // 复位上升沿清故障锁存 [-] / reset rising edge clears the fault latch
    bStepStart     : BOOL := FALSE;          // 阶跃施加时刻的上升沿（调用方给出）[-] / rising edge at the step application instant
    fMvStep        : REAL := 10.0;           // 操纵量阶跃幅度（带符号）[工程单位] / manipulated variable step amplitude, signed [engineering unit]
    fMvStepEps     : REAL := 1.0E-3;         // 阶跃幅度可辨下限 [工程单位] / step amplitude recognisable floor [engineering unit]
    fPv            : REAL := 0.0;            // 过程量实测 [工程单位] / measured process variable [engineering unit]
    fSampleS       : REAL := 0.1;            // 采样拍周期 [秒]，域 1E-4..10 / sample period [second], domain 1E-4 to 10
    tTimeout       : TIME := T#300S;         // 上升相超时 [毫秒] / rise phase timeout [millisecond]
    tSettle        : TIME := T#5S;           // 稳定确认时长 [毫秒] / settle confirmation duration [millisecond]
    fSettleBandPct : REAL := 1.0;            // 稳定带，占当前跨度百分比 [百分比] / settle band as a percentage of the current span [percent]
    fMinDeltaPv    : REAL := 0.5;            // 响应最小可辨量 [工程单位] / minimum recognisable response [engineering unit]
    bUseTangent    : BOOL := FALSE;          // 真 = 出口取切线法，假 = 出口取两点法 [-] / true selects the tangent method, false selects the two-point method
    fTauMinS       : REAL := 0.2;            // 时间常数可接受下限 [秒] / acceptable time constant floor [second]
    fTauMaxS       : REAL := 7200.0;         // 时间常数可接受上限 [秒] / acceptable time constant ceiling [second]
    fDeadMaxS      : REAL := 600.0;          // 纯延迟可接受上限 [秒] / acceptable dead time ceiling [second]
END_VAR
VAR_OUTPUT
    fGainK         : REAL := 0.0;            // 辨识增益 K [工程单位比] / identified process gain [engineering unit ratio]
    fTauS          : REAL := 0.0;            // 辨识时间常数 T [秒] / identified time constant [second]
    fDeadS         : REAL := 0.0;            // 辨识纯延迟 L [秒] / identified dead time [second]
    fDeltaPv       : REAL := 0.0;            // 本次阶跃的总过程量变化 [工程单位] / total process change of this step [engineering unit]
    fPvBase        : REAL := 0.0;            // 阶跃前基线过程量 [工程单位] / baseline process variable before the step [engineering unit]
    fPvFinal       : REAL := 0.0;            // 稳定后过程量 [工程单位] / settled process variable [engineering unit]
    fTauTwoPointS  : REAL := 0.0;            // 两点法时间常数 [秒] / two-point method time constant [second]
    fDeadTwoPointS : REAL := 0.0;            // 两点法纯延迟 [秒] / two-point method dead time [second]
    fTauTangentS   : REAL := 0.0;            // 切线法时间常数 [秒] / tangent method time constant [second]
    fDeadTangentS  : REAL := 0.0;            // 切线法纯延迟 [秒] / tangent method dead time [second]
    bValid         : BOOL := FALSE;          // 参数是否可交付 [-] / parameters deliverable flag
    bIdentDone     : BOOL := FALSE;          // 辨识完成单拍脉冲 [-] / identification done single-shot pulse
    eState         : E_DL_FopdtState := E_DL_FopdtState.eIdle; // 相位出口，段尾单点映射 [枚举] / phase outlet, single-point mapped at the tail
    eCause         : E_DL_FopdtCause := E_DL_FopdtCause.eNone; // 成因出口，锁存至复位 [枚举] / cause outlet, latched until reset
    bError         : BOOL := FALSE;          // 故障锁存标志 [-] / fault latch flag
END_VAR
VAR
    rtStep         : R_TRIG;                 // 阶跃沿检测，段 0 无条件刷新 / step edge detector, refreshed unconditionally in segment zero
    rtReset        : R_TRIG;                 // 复位沿检测，段 0 无条件刷新 / reset edge detector, refreshed unconditionally in segment zero
    tonTimeout     : TON;                    // 上升相超时计时，段 0 无条件刷新 / rise phase timeout timer, refreshed unconditionally in segment zero
    tonSettle      : TON;                    // 稳定确认计时，段 0 无条件刷新 / settle confirmation timer, refreshed unconditionally in segment zero
    _eState        : E_DL_FopdtState := E_DL_FopdtState.eIdle;  // 内部相位，CASE 唯一写入目标 / internal phase, the only CASE write target
    _eCause        : E_DL_FopdtCause := E_DL_FopdtCause.eNone;  // 内部成因，锁存量 / internal cause, latched quantity
    _bFault        : BOOL := FALSE;          // 故障锁存位 [-] / fault latch bit
    _bValid        : BOOL := FALSE;          // 参数有效内部位，锁存至下次辨识 / internal validity bit, latched until the next identification
    _bIdentInt     : BOOL := FALSE;          // 完成脉冲内部位，统一出口映射 / internal done bit, mapped at the unified outlet
    _bInit         : BOOL := FALSE;          // 首扫初始化完成标志（R310）/ first scan initialisation flag
    _bSampleOk     : BOOL := FALSE;          // 本拍样本有效（过程量有限）[-] / this-scan sample valid flag
    _bStoreOk      : BOOL := FALSE;          // 环窗槽位合法可写 [-] / ring slot legal and writable
    _bSpanOk       : BOOL := FALSE;          // 跨度估计可用于稳定带判据 [-] / span estimate usable for the settle band
    _bCfgBad       : BOOL := FALSE;          // 组态非法标志 [-] / illegal configuration flag
    _bCross28      : BOOL := FALSE;          // 已捕获 28.3% 穿越点 [-] / 28.3 percent crossing captured
    _bCross63      : BOOL := FALSE;          // 已捕获 63.2% 穿越点 [-] / 63.2 percent crossing captured
    _bDeadClamped  : BOOL := FALSE;          // 纯延迟负值已按零处理 [-] / negative dead time forced to zero
    _nHead         : INT := 0;               // 环窗最近样本槽位（1 起，回钳 1..N）[槽号] / newest ring slot, one-based, clamped one through N
    _nFill         : INT := 0;               // 环窗已填样本数（0..N）[个] / samples held in the ring [count]
    _nIdx          : INT := 0;               // 环窗下标游标 [槽号] / ring index cursor [slot]
    _nPrev         : INT := 0;               // 时间序前一槽位 [槽号] / previous slot in time order [slot]
    _nGuard        : INT := 0;               // 遍历防死循环守护计数 [次] / traversal guard against runaway loops [count]
    _nK            : INT := 0;               // 时间序遍历序号（1 = 最旧样本）[序号] / time-order ordinal, one is the oldest [ordinal]
    _fDtS          : REAL := 0.1;            // 钳定后的采样拍周期 [秒] / clamped sample period [second]
    _fElapsedS     : REAL := 0.0;            // 上升相已历时 [秒] / elapsed time within the rise phase [second]
    _fPvPrev       : REAL := 0.0;            // 上一拍过程量快照 [工程单位] / previous scan process value snapshot [engineering unit]
    _fPvBase       : REAL := 0.0;            // 基线过程量（时间序最旧样本）[工程单位] / baseline process value from the oldest sample [engineering unit]
    _fPvNow        : REAL := 0.0;            // 本拍样本过程量 [工程单位] / current sample process value [engineering unit]
    _fPvFinal      : REAL := 0.0;            // 稳定后过程量（时间序最新样本）[工程单位] / settled process value from the newest sample [engineering unit]
    _fPvOld        : REAL := 0.0;            // 遍历中的前一有效样本过程量 [工程单位] / previous valid sample during traversal [engineering unit]
    _fDeltaPv      : REAL := 0.0;            // 总过程量变化 [工程单位] / total process change [engineering unit]
    _fSpan         : REAL := 0.0;            // 已观测过程量跨度上确界 [工程单位] / supremum of the observed process span [engineering unit]
    _fSettleAbs    : REAL := 0.0;            // 稳定带绝对量 [工程单位] / absolute settle band [engineering unit]
    _fFrac         : REAL := 0.0;            // 归一化响应分数（0..1）[无量纲] / normalised response fraction [dimensionless]
    _fSlopeNow     : REAL := 0.0;            // 本拍斜率 [工程单位每秒] / slope of this scan [engineering unit per second]
    _fSlopeMax     : REAL := 0.0;            // 最大斜率上确界 [工程单位每秒] / supremum of the slope magnitude [engineering unit per second]
    _fSlopeSig     : REAL := 0.0;            // 带符号最大斜率，符号取 SIGN(ΔPV) [工程单位每秒] / signed maximum slope carrying the delta PV sign [engineering unit per second]
    _fSlopeLoc     : REAL := 0.0;            // 相邻样本斜率 [工程单位每秒] / slope between adjacent samples [engineering unit per second]
    _fDtLoc        : REAL := 0.0;            // 相邻样本时差 [秒] / time difference between adjacent samples [second]
    _fT28          : REAL := 0.0;            // 28.3% 穿越时刻 [秒] / 28.3 percent crossing instant [second]
    _fT63          : REAL := 0.0;            // 63.2% 穿越时刻 [秒] / 63.2 percent crossing instant [second]
    _fTSlopeMax    : REAL := 0.0;            // 最大斜率出现时刻 [秒] / instant of the maximum slope [second]
    _fPvSlopeMax   : REAL := 0.0;            // 最大斜率处过程量 [工程单位] / process value at the maximum slope [engineering unit]
    _fTauTwo       : REAL := 0.0;            // 两点法时间常数计算值 [秒] / two-point time constant, computed value [second]
    _fDeadTwo      : REAL := 0.0;            // 两点法纯延迟计算值 [秒] / two-point dead time, computed value [second]
    _fTauTan       : REAL := 0.0;            // 切线法时间常数计算值 [秒] / tangent time constant, computed value [second]
    _fDeadTan      : REAL := 0.0;            // 切线法纯延迟计算值 [秒] / tangent dead time, computed value [second]
    _fTauOut       : REAL := 0.0;            // 出口选用时间常数 [秒] / selected outlet time constant [second]
    _fDeadOut      : REAL := 0.0;            // 出口选用纯延迟 [秒] / selected outlet dead time [second]
    _fGain         : REAL := 0.0;            // 增益计算值 [工程单位比] / computed gain [engineering unit ratio]
    _fMvDen        : REAL := 0.0;            // 增益分母（阶跃幅度）暂存 [工程单位] / gain denominator held in a local [engineering unit]
    _fGainK        : REAL := 0.0;            // 出口保持：增益 [工程单位比] / outlet holder for the gain [engineering unit ratio]
    _fTauS         : REAL := 0.0;            // 出口保持：时间常数 [秒] / outlet holder for the time constant [second]
    _fDeadS        : REAL := 0.0;            // 出口保持：纯延迟 [秒] / outlet holder for the dead time [second]
    _fDeltaPvOut   : REAL := 0.0;            // 出口保持：总变化量 [工程单位] / outlet holder for the total change [engineering unit]
    _fPvBaseOut    : REAL := 0.0;            // 出口保持：基线过程量 [工程单位] / outlet holder for the baseline value [engineering unit]
    _fPvFinalOut   : REAL := 0.0;            // 出口保持：稳定点过程量 [工程单位] / outlet holder for the settled value [engineering unit]
    _fTauTwoOut    : REAL := 0.0;            // 出口保持：两点法时间常数 [秒] / outlet holder for the two-point time constant [second]
    _fDeadTwoOut   : REAL := 0.0;            // 出口保持：两点法纯延迟 [秒] / outlet holder for the two-point dead time [second]
    _fTauTanOut    : REAL := 0.0;            // 出口保持：切线法时间常数 [秒] / outlet holder for the tangent time constant [second]
    _fDeadTanOut   : REAL := 0.0;            // 出口保持：切线法纯延迟 [秒] / outlet holder for the tangent dead time [second]
    _afPvV         : ARRAY[1..512] OF REAL := [512(0.0)]; // 环窗过程量缓存 [工程单位] / ring buffer of process values [engineering unit]
    _afPvT         : ARRAY[1..512] OF REAL := [512(0.0)]; // 环窗时刻缓存，与过程量同槽同步写入 [秒] / ring buffer of instants, lockstep with the values [second]
END_VAR
VAR CONSTANT
    DL_FOPDT_MAX    : INT := 512;            // 环窗容量与槽位回钳上界 [个] / ring capacity and slot clamp upper bound [count]
    DL_FOPDT_SMIN   : REAL := 1.0E-4;        // 采样周期下限，防除零 [秒] / sample period floor against division by zero [second]
    DL_FOPDT_SMAX   : REAL := 10.0;          // 采样周期上限，防时基错配 [秒] / sample period ceiling against a mismatched time base [second]
    DL_FOPDT_DTMIN  : REAL := 1.0E-6;        // 相邻样本时差下限，斜率除子 [秒] / adjacent sample time difference floor for the slope divisor [second]
    DL_FOPDT_FRAC28 : REAL := 0.283;         // 两点法第一穿越点 [无量纲] / two-point first crossing fraction [dimensionless]
    DL_FOPDT_FRAC63 : REAL := 0.632;         // 两点法第二穿越点 [无量纲] / two-point second crossing fraction [dimensionless]
    DL_FOPDT_TAUCOEF: REAL := 1.5;           // 两点法时间常数系数 [无量纲] / two-point time constant coefficient [dimensionless]
    DL_FOPDT_EPS    : REAL := 1.0E-9;        // 斜率与分数类除子下限 [无量纲] / floor for slope and fraction divisors [dimensionless]
    DL_FOPDT_GAINMAX: REAL := 1.0E9;         // 增益量级上限，防量纲错配 [工程单位比] / gain magnitude ceiling against a dimension mismatch [engineering unit ratio]
    DL_FOPDT_GUARD  : INT := 1024;           // 遍历守护上限，两倍容量 [次] / traversal guard, twice the capacity [count]
    DL_FOPDT_MINPTS : INT := 4;              // 参与辨识的最少样本数 [个] / minimum sample count for identification [count]
END_VAR

// 段 0｜定时器与沿检测无条件周期刷新（禁入分支），IN 只串状态闸 / segment 0, unconditional refresh of timers and edge detectors with state gates on IN only
rtStep(CLK := bStepStart); // 阶跃沿检测无条件刷新 / unconditional refresh of the step edge detector
rtReset(CLK := bReset); // 复位沿检测无条件刷新 / unconditional refresh of the reset edge detector
tonTimeout(IN := (_eState = E_DL_FopdtState.eRise) AND (NOT _bFault), PT := tTimeout); // 上升相超时，IN 串相位闸与故障闸 / rise phase timeout, IN carries the phase gate and the fault gate
tonSettle(IN := (_eState = E_DL_FopdtState.eRise) AND _bSampleOk AND _bSpanOk AND (ABS(fPv - _fPvPrev) <= _fSettleAbs), PT := tSettle); // 稳定确认，IN 串相位闸与稳定带判据 / settle confirmation with the phase gate and the settle band criterion on IN

// 段 1｜首扫初始化（R310）：学习量与环窗从确定起点开始 / segment 1, first scan initialisation so that learning quantities and the ring start known
IF NOT _bInit THEN // 首扫一拍 / the very first scan
    _bInit := TRUE; // 置首扫完成标志 / raise the first scan flag
    _eState := E_DL_FopdtState.eIdle; // 相位从空闲起步 / the phase starts from idle
    _eCause := E_DL_FopdtCause.eNone; // 成因清零 / clear the cause
    _bFault := FALSE; // 故障锁存清零 / clear the fault latch
    _bValid := FALSE; // 有效位清零 / clear the validity bit
    _nHead := 0; // 环窗无样本 / the ring holds no sample
    _nFill := 0; // 环窗计数清零 / clear the ring count
    _fSpan := 0.0; // 跨度估计清零 / clear the span estimate
END_IF

// 段 2｜复位沿作用域逐项声明：清锁存 / 迁相位 / 清累计量 / segment 2, reset edge scope declared item by item
IF rtReset.Q OR (NOT bEnable) THEN // 复位沿或失能 / reset edge or disabled
    _bFault := FALSE; // 作用域一：清故障锁存 / scope one, clear the fault latch
    _eCause := E_DL_FopdtCause.eNone; // 作用域一：清成因 / scope one, clear the cause
    _bIdentInt := FALSE; // 作用域一：清完成脉冲内部位 / scope one, clear the internal done bit
    _eState := E_DL_FopdtState.eIdle; // 作用域二：迁回空闲相 / scope two, migrate back to idle
    _nHead := 0; // 作用域三：清环窗槽位 / scope three, clear the ring slot cursor
    _nFill := 0; // 作用域三：清环窗计数 / scope three, clear the ring count
    _fSpan := 0.0; // 作用域三：清跨度估计 / scope three, clear the span estimate
    _fElapsedS := 0.0; // 作用域三：清历时 / scope three, clear the elapsed time
END_IF

// 段 3｜组态域闸（R151）：参与判据换算的每个引脚逐项闸，缺一即判据静默失效 / segment 3, configuration domain gate over every pin used by the criteria
_bCfgBad := FALSE; // 组态非法标志预置假 / preset the illegal configuration flag to false
IF (fSampleS <> fSampleS) THEN // 采样周期 NaN 自反判 / NaN detection on the sample period
    _bCfgBad := TRUE; // 判组态非法 / illegal configuration
END_IF
IF (fSampleS < DL_FOPDT_SMIN) OR (fSampleS > DL_FOPDT_SMAX) THEN // 采样周期越域 / sample period out of domain
    _bCfgBad := TRUE; // 判组态非法 / illegal configuration
END_IF
IF (fMvStep <> fMvStep) OR ((fMvStep - fMvStep) <> (fMvStep - fMvStep)) THEN // 阶跃幅度非有限 / step amplitude non-finite
    _bCfgBad := TRUE; // 判组态非法 / illegal configuration
END_IF
IF (fMvStepEps <= 0.0) OR (fMvStepEps <> fMvStepEps) THEN // 幅度可辨下限非正或非有限 / amplitude floor not positive or non-finite
    _bCfgBad := TRUE; // 判组态非法 / illegal configuration
END_IF
IF (fMinDeltaPv <= 0.0) OR (fMinDeltaPv <> fMinDeltaPv) THEN // 最小可辨量非正或非有限 / response floor not positive or non-finite
    _bCfgBad := TRUE; // 判组态非法 / illegal configuration
END_IF
IF (fSettleBandPct <= 0.0) OR (fSettleBandPct >= 100.0) OR (fSettleBandPct <> fSettleBandPct) THEN // 稳定带百分比越域 / settle band percentage out of domain
    _bCfgBad := TRUE; // 判组态非法 / illegal configuration
END_IF
IF (fTauMinS <= 0.0) OR (fTauMaxS <= fTauMinS) OR (fTauMaxS <> fTauMaxS) THEN // 时间常数上下限自相矛盾 / time constant bounds contradict each other
    _bCfgBad := TRUE; // 判组态非法 / illegal configuration
END_IF
IF (fDeadMaxS < 0.0) OR (fDeadMaxS <> fDeadMaxS) THEN // 纯延迟上限为负或非有限 / dead time ceiling negative or non-finite
    _bCfgBad := TRUE; // 判组态非法 / illegal configuration
END_IF
IF (tTimeout <= T#0S) OR (tSettle <= T#0S) THEN // 时间引脚非正 / time pins not positive
    _bCfgBad := TRUE; // 判组态非法 / illegal configuration
END_IF
IF tSettle >= tTimeout THEN // 稳定窗不短于相超时窗，违反双窗配比（R100）/ the settle window is not shorter than the phase timeout
    _bCfgBad := TRUE; // 判组态非法 / illegal configuration
END_IF
IF _bCfgBad AND (NOT _bFault) THEN // 组态非法且未锁存 / illegal configuration and not yet latched
    _eCause := E_DL_FopdtCause.eCfgIllegal; // 成因记组态非法 / record the illegal configuration cause
    _bFault := TRUE; // 置故障锁存 / raise the fault latch
    _bValid := FALSE; // 参数不可交付 / parameters not deliverable
    _eState := E_DL_FopdtState.eFault; // 迁故障相 / migrate to the fault phase
END_IF

// 段 4｜本拍量预置（单拍标志限域，不含快照与环窗保持量）/ segment 4, per-scan presets limited to single-shot flags
_fDtS := fSampleS; // 采样周期直通 / sample period passes through
IF _fDtS < DL_FOPDT_SMIN THEN // 周期过小 / period too small
    _fDtS := DL_FOPDT_SMIN; // 抬到下限，防时基除零 / raised against a zero time base
ELSIF _fDtS > DL_FOPDT_SMAX THEN // 周期过大 / period too large
    _fDtS := DL_FOPDT_SMAX; // 压到上限 / pressed to the ceiling
END_IF
_bSampleOk := (fPv = fPv) AND ((fPv - fPv) = (fPv - fPv)); // 过程量有限性闸，NaN 用自反、无穷用差值自减 / process value finiteness gate
_fPvNow := fPv; // 本拍样本默认取实测 / the current sample defaults to the measurement
IF NOT _bSampleOk THEN // 非有限拍 / non-finite scan
    _fPvNow := _fPvPrev; // 非有限不穿透：改取上拍快照 / nothing non-finite passes, the previous snapshot is used
END_IF
_fSettleAbs := _fSpan * fSettleBandPct / 100.0; // 稳定带绝对量，除子为常量 100.0 / absolute settle band, the divisor is the literal constant one hundred
_bSpanOk := _fSpan > 0.0; // 跨度估计可用性 / span estimate availability

// 段 5｜相位机：ENUM + CASE，含 ELSE 非法相位兜底（R128）/ segment 5, phase machine with an ELSE fallback for illegal phases
CASE _eState OF
E_DL_FopdtState.eIdle: // 空闲相：等阶跃上升沿 / idle phase, waiting for the step rising edge
    IF rtStep.Q THEN // 阶跃沿到达 / the step edge arrived
        _nHead := 0; // 环窗槽位清零 / clear the ring slot cursor
        _nFill := 0; // 环窗计数清零 / clear the ring count
        _fSpan := 0.0; // 跨度估计清零 / clear the span estimate
        _fElapsedS := 0.0; // 历时清零 / clear the elapsed time
        _fSlopeMax := 0.0; // 最大斜率清零 / clear the maximum slope
        _fPvSlopeMax := 0.0; // 最大斜率处过程量清零 / clear the value at the maximum slope
        _fTSlopeMax := 0.0; // 最大斜率时刻清零 / clear the instant of the maximum slope
        _bCross28 := FALSE; // 穿越标志清零 / clear the crossing flag
        _bCross63 := FALSE; // 穿越标志清零 / clear the crossing flag
        _fPvPrev := fPv; // 基线快照取当拍实测 / the baseline snapshot takes the current measurement
        _fPvBase := fPv; // 基线过程量取当拍实测 / the baseline process value takes the current measurement
        _eState := E_DL_FopdtState.eRise; // 迁上升相 / migrate to the rise phase
    END_IF

E_DL_FopdtState.eRise: // 上升相：缓存样本、跟踪斜率与跨度 / rise phase, buffering samples and tracking slope and span
    _fElapsedS := _fElapsedS + _fDtS; // 累计历时 / accumulate the elapsed time
    _bStoreOk := FALSE; // 写入许可预置假 / preset the write permit to false
    IF _nFill < DL_FOPDT_MAX THEN // 环窗未满 / the ring is not yet full
        _nHead := _nHead + 1; // 槽位前移，天然落在 1..N / advance the slot, naturally inside one through N
        _nFill := _nFill + 1; // 计数递增 / increment the count
        _bStoreOk := TRUE; // 允许写入 / writing permitted
    ELSE // 环窗已满 / the ring is full
        _nHead := _nHead + 1; // 槽位前移 / advance the slot
        IF _nHead > DL_FOPDT_MAX THEN // 越过上界 / past the upper bound
            _nHead := 1; // 回钳到一号槽（环窗回钳口径）/ clamp back to slot one
        END_IF
        _bStoreOk := TRUE; // 允许写入 / writing permitted
    END_IF
    IF _bStoreOk THEN // 槽位合法 / slot is legal
        _afPvV[_nHead] := _fPvNow; // 过程量入环窗 / store the process value
        _afPvT[_nHead] := _fElapsedS; // 时刻同步入同槽 / store the instant into the same slot
    END_IF
    IF ABS(_fPvNow - _fPvBase) > _fSpan THEN // 跨度取绝对偏差上确界 / the span takes the supremum of absolute deviation
        _fSpan := ABS(_fPvNow - _fPvBase); // 更新跨度 / refresh the span
    END_IF
    _fSlopeNow := ABS(_fPvNow - _fPvPrev) / _fDtS; // 本拍斜率绝对值，除子已钳定大于零 / absolute slope of this scan, divisor proven positive
    IF _fSlopeNow > _fSlopeMax THEN // 斜率上确界跟踪 / supremum slope tracking
        _fSlopeMax := _fSlopeNow; // 更新最大斜率 / refresh the maximum slope
        _fPvSlopeMax := _fPvNow; // 记录该点过程量 / record the value at that point
        _fTSlopeMax := _fElapsedS; // 记录该点时刻 / record the instant of that point
    END_IF
    _fPvPrev := _fPvNow; // 快照推进 / advance the snapshot
    IF tonSettle.Q OR tonTimeout.Q THEN // 稳定达成或超时 / settled or timed out
        _eState := E_DL_FopdtState.eEval; // 迁评估相 / migrate to the evaluation phase
    END_IF

E_DL_FopdtState.eEval: // 评估相：按时间序遍历环窗，两法并行求解 / evaluation phase, traversal in time order with both methods solved
    _nK := _nFill; // 参与判定的样本数 / samples participating in the verdict
    IF _nK > DL_FOPDT_MAX THEN // 防御：计数不得越容 / defence, the count must not exceed capacity
        _nK := DL_FOPDT_MAX; // 回钳到容量 / clamp to the capacity
    END_IF
    IF _nK < DL_FOPDT_MINPTS THEN // 样本不足 / too few samples
        _eCause := E_DL_FopdtCause.eNoCross; // 成因记样本不足缺穿越点 / record the missing crossing cause
        _bFault := TRUE; // 置故障锁存 / raise the fault latch
        _bValid := FALSE; // 参数不可交付 / parameters not deliverable
        _eState := E_DL_FopdtState.eFault; // 迁故障相 / migrate to the fault phase
    ELSE
        _nIdx := _nHead - _nFill + 1; // 时间序最旧槽位 / the oldest slot in time order
        IF _nIdx < 1 THEN // 越过下界 / below the lower bound
            _nIdx := _nIdx + DL_FOPDT_MAX; // 单次回绕补齐（时间序回钳）/ a single wrap restores the time order
        END_IF
        _fPvBase := _afPvV[_nIdx]; // 基线取时间序最旧样本 / the baseline takes the oldest sample
        _fPvOld := _fPvBase; // 遍历起点过程量 / traversal start value
        _fPvFinal := _afPvV[_nHead]; // 稳定点取时间序最新样本 / the settled value takes the newest sample
        _fDeltaPv := _fPvFinal - _fPvBase; // 总变化量 / total change
        IF ABS(_fDeltaPv) <= fMinDeltaPv THEN // 响应不足 / response too small
            _eCause := E_DL_FopdtCause.eLackResp; // 成因记响应不足 / record the insufficient response cause
            _bFault := TRUE; // 置故障锁存 / raise the fault latch
            _bValid := FALSE; // 参数不可交付 / parameters not deliverable
            _eState := E_DL_FopdtState.eFault; // 迁故障相 / migrate to the fault phase
        ELSIF ABS(fMvStep) <= fMvStepEps THEN // 阶跃幅度近零 / step amplitude near zero
            _eCause := E_DL_FopdtCause.eMvZero; // 成因记幅度近零 / record the near-zero amplitude cause
            _bFault := TRUE; // 置故障锁存 / raise the fault latch
            _bValid := FALSE; // 参数不可交付 / parameters not deliverable
            _eState := E_DL_FopdtState.eFault; // 迁故障相 / migrate to the fault phase
        ELSE
            _bCross28 := FALSE; // 穿越标志复位 / clear the crossing flag
            _bCross63 := FALSE; // 穿越标志复位 / clear the crossing flag
            _nGuard := 0; // 遍历守护计数清零 / reset the traversal guard
            _nK := 1; // 自最旧样本起按时间序遍历（R194）/ traverse from the oldest sample in time order
            WHILE (_nK <= _nFill) AND (_nGuard < DL_FOPDT_GUARD) DO // 双重守护：样本数与计数上限 / dual guard on the sample count and the counter cap
                _nGuard := _nGuard + 1; // 守护计数递增 / increment the guard
                _nIdx := _nHead - _nFill + _nK; // 时间序槽位 / the slot in time order
                IF _nIdx < 1 THEN // 越过下界 / below the lower bound
                    _nIdx := _nIdx + DL_FOPDT_MAX; // 单次回绕 / single wrap
                END_IF
                _fFrac := (_afPvV[_nIdx] - _fPvBase) / _fDeltaPv; // 归一化响应分数，除子绝对值已证超可辨量 / normalised fraction, divisor proven above the floor
                IF (NOT _bCross28) AND (_fFrac >= DL_FOPDT_FRAC28) THEN // 首次越过 28.3% / first crossing of 28.3 percent
                    _fT28 := _afPvT[_nIdx]; // 记录穿越时刻 / record the crossing instant
                    _bCross28 := TRUE; // 置穿越标志 / raise the crossing flag
                END_IF
                IF (NOT _bCross63) AND (_fFrac >= DL_FOPDT_FRAC63) THEN // 首次越过 63.2% / first crossing of 63.2 percent
                    _fT63 := _afPvT[_nIdx]; // 记录穿越时刻 / record the crossing instant
                    _bCross63 := TRUE; // 置穿越标志 / raise the crossing flag
                END_IF
                IF _nK > 1 THEN // 自第二个样本起可算斜率 / slopes exist from the second sample onward
                    _nPrev := _nIdx - 1; // 前一槽位 / the previous slot
                    IF _nPrev < 1 THEN // 越过下界 / below the lower bound
                        _nPrev := _nPrev + DL_FOPDT_MAX; // 单次回绕 / single wrap
                    END_IF
                    _fDtLoc := _afPvT[_nIdx] - _afPvT[_nPrev]; // 相邻样本时差 / adjacent sample time difference
                    IF _fDtLoc > DL_FOPDT_DTMIN THEN // 时差可用 / the difference is usable
                        _fSlopeLoc := ABS((_afPvV[_nIdx] - _fPvOld) / _fDtLoc); // 局部斜率绝对值 / local absolute slope
                        IF _fSlopeLoc > _fSlopeMax THEN // 斜率上确界 / slope supremum
                            _fSlopeMax := _fSlopeLoc; // 更新最大斜率 / refresh the maximum slope
                            _fPvSlopeMax := _afPvV[_nIdx]; // 记录该点过程量 / record the value at that point
                            _fTSlopeMax := _afPvT[_nIdx]; // 记录该点时刻 / record the instant of that point
                        END_IF
                    END_IF
                END_IF
                _fPvOld := _afPvV[_nIdx]; // 推进前一有效样本 / advance the previous valid sample
                _nK := _nK + 1; // 序号递增 / increment the ordinal
            END_WHILE
            IF (NOT _bCross28) OR (NOT _bCross63) THEN // 缺穿越点 / a crossing is missing
                _eCause := E_DL_FopdtCause.eNoCross; // 成因记缺穿越点 / record the missing crossing cause
                _bFault := TRUE; // 置故障锁存 / raise the fault latch
                _bValid := FALSE; // 参数不可交付 / parameters not deliverable
                _eState := E_DL_FopdtState.eFault; // 迁故障相 / migrate to the fault phase
            ELSIF (_fT63 - _fT28) < DL_FOPDT_DTMIN THEN // 两穿越点重合，时间常数不可辨 / the crossings coincide and the time constant is unresolvable
                _eCause := E_DL_FopdtCause.eNoCross; // 成因记穿越点不可辨 / record the unresolvable crossing cause
                _bFault := TRUE; // 置故障锁存 / raise the fault latch
                _bValid := FALSE; // 参数不可交付 / parameters not deliverable
                _eState := E_DL_FopdtState.eFault; // 迁故障相 / migrate to the fault phase
            ELSE
                _fTauTwo := DL_FOPDT_TAUCOEF * (_fT63 - _fT28); // 两点法时间常数 / two-point time constant
                _fDeadTwo := _fT63 - _fTauTwo; // 两点法纯延迟 / two-point dead time
                _bDeadClamped := FALSE; // 钳位标志复位 / clear the clamp flag
                IF _fDeadTwo < 0.0 THEN // 延迟负值不可能 / a negative dead time is impossible
                    _fDeadTwo := 0.0; // 按零处理 / forced to zero
                    _bDeadClamped := TRUE; // 置钳位标志 / raise the clamp flag
                END_IF
                IF _fSlopeMax > DL_FOPDT_EPS THEN // 斜率可用 / the slope is usable
                    _fSlopeSig := _fSlopeMax * SIGN(_fDeltaPv); // 带符号斜率：SIGN(ΔPV) ∈ {-1, 1}（ΔPV 已证 |·| > fMinDeltaPv > 0），量级仍由 _fSlopeMax 超阈证明 / signed slope, the sign of delta PV is proven nonzero and the magnitude stays proven by the slope floor
                    _fTauTan := _fDeltaPv / _fSlopeSig; // 切线法时间常数，除子量级已证超阈且符号与分子同源 / tangent time constant, the divisor magnitude is proven and its sign matches the numerator
                    _fDeadTan := _fTSlopeMax - (_fPvSlopeMax - _fPvBase) / _fSlopeSig; // 切线法纯延迟：截距用带符号斜率，负向阶跃不再系统性高估（R56 返修）/ tangent dead time, the intercept uses the signed slope so a negative step no longer overestimates
                    IF _fDeadTan < 0.0 THEN // 延迟负值不可能 / a negative dead time is impossible
                        _fDeadTan := 0.0; // 按零处理 / forced to zero
                        _bDeadClamped := TRUE; // 置钳位标志 / raise the clamp flag
                    END_IF
                ELSE // 斜率不可用 / the slope is unusable
                    _fTauTan := _fTauTwo; // 以两点法兜底 / fall back to the two-point result
                    _fDeadTan := _fDeadTwo; // 纯延迟同款兜底 / the dead time falls back the same way
                END_IF
                _fMvDen := fMvStep; // 增益分母落局部量 / the gain denominator lands in a local
                IF ABS(_fMvDen) <= fMvStepEps THEN // 分母近零 / denominator near zero
                    _eCause := E_DL_FopdtCause.eMvZero; // 成因记幅度近零 / record the near-zero amplitude cause
                    _bFault := TRUE; // 置故障锁存 / raise the fault latch
                    _bValid := FALSE; // 参数不可交付 / parameters not deliverable
                    _eState := E_DL_FopdtState.eFault; // 迁故障相 / migrate to the fault phase
                ELSE
                    _fGain := _fDeltaPv / _fMvDen; // 增益 = ΔPV / ΔMV / gain equals delta PV over delta MV
                    IF ABS(_fGain) > DL_FOPDT_GAINMAX THEN // 增益量级越界 / gain magnitude out of range
                        _eCause := E_DL_FopdtCause.eCfgIllegal; // 成因记组态非法（量纲错配）/ record illegal configuration, dimension mismatch
                        _bFault := TRUE; // 置故障锁存 / raise the fault latch
                        _bValid := FALSE; // 参数不可交付 / parameters not deliverable
                        _eState := E_DL_FopdtState.eFault; // 迁故障相 / migrate to the fault phase
                    ELSE
                        _fTauOut := _fTauTwo; // 出口时间常数默认取两点法 / the outlet time constant defaults to the two-point result
                        _fDeadOut := _fDeadTwo; // 出口纯延迟默认取两点法 / the outlet dead time defaults to the two-point result
                        IF bUseTangent THEN // 切线法优先 / the tangent method takes precedence
                            _fTauOut := _fTauTan; // 取切线法时间常数 / take the tangent time constant
                            _fDeadOut := _fDeadTan; // 取切线法纯延迟 / take the tangent dead time
                        END_IF
                        IF (_fTauOut < fTauMinS) OR (_fTauOut > fTauMaxS) THEN // 时间常数越接受域 / time constant outside the acceptable domain
                            _eCause := E_DL_FopdtCause.eCfgIllegal; // 成因记组态非法（接受域不匹配）/ record illegal configuration, bound mismatch
                            _bFault := TRUE; // 置故障锁存 / raise the fault latch
                            _bValid := FALSE; // 参数不可交付 / parameters not deliverable
                            _eState := E_DL_FopdtState.eFault; // 迁故障相 / migrate to the fault phase
                        ELSIF _fDeadOut > fDeadMaxS THEN // 纯延迟越接受域 / dead time outside the acceptable domain
                            _eCause := E_DL_FopdtCause.eCfgIllegal; // 成因记组态非法（接受域不匹配）/ record illegal configuration, bound mismatch
                            _bFault := TRUE; // 置故障锁存 / raise the fault latch
                            _bValid := FALSE; // 参数不可交付 / parameters not deliverable
                            _eState := E_DL_FopdtState.eFault; // 迁故障相 / migrate to the fault phase
                        ELSE
                            _fGainK := _fGain; // 增益落定 / settle the gain
                            _fTauS := _fTauOut; // 时间常数落定 / settle the time constant
                            _fDeadS := _fDeadOut; // 纯延迟落定 / settle the dead time
                            _fDeltaPvOut := _fDeltaPv; // 总变化量落定 / settle the total change
                            _fTauTwoOut := _fTauTwo; // 两点法时间常数落定 / settle the two-point time constant
                            _fDeadTwoOut := _fDeadTwo; // 两点法纯延迟落定 / settle the two-point dead time
                            _fTauTanOut := _fTauTan; // 切线法时间常数落定 / settle the tangent time constant
                            _fDeadTanOut := _fDeadTan; // 切线法纯延迟落定 / settle the tangent dead time
                            _fPvBaseOut := _fPvBase; // 基线落定 / settle the baseline
                            _fPvFinalOut := _fPvFinal; // 稳定点落定 / settle the settled value
                            _bValid := TRUE; // 参数可交付（锁存至下一次辨识）/ parameters deliverable until the next identification
                            _bIdentInt := TRUE; // 完成脉冲内部位置位（统一出口映射，R187）/ raise the internal done bit, mapped at the unified outlet
                            IF _bDeadClamped THEN // 延迟负值已钳零 / the dead time was clamped to zero
                                _eCause := E_DL_FopdtCause.eDeadNeg; // 信息级成因，不置故障标志 / informational cause without raising the fault flag
                            END_IF
                            _eState := E_DL_FopdtState.eDone; // 迁完成相 / migrate to the done phase
                        END_IF
                    END_IF
                END_IF
            END_IF
        END_IF
    END_IF

E_DL_FopdtState.eDone: // 完成相：参数驻留，仅接受复位或新阶跃 / done phase, parameters held, only reset or a new step accepted
    IF rtStep.Q THEN // 新阶跃沿 / a new step edge
        _nHead := 0; // 环窗槽位清零 / clear the ring slot cursor
        _nFill := 0; // 环窗计数清零 / clear the ring count
        _fSpan := 0.0; // 跨度估计清零 / clear the span estimate
        _fElapsedS := 0.0; // 历时清零 / clear the elapsed time
        _fSlopeMax := 0.0; // 最大斜率清零 / clear the maximum slope
        _fPvSlopeMax := 0.0; // 最大斜率处过程量清零（R56 返修补齐，与空闲相分支对齐）/ clear the value at the maximum slope, aligned with the idle branch
        _fTSlopeMax := 0.0; // 最大斜率时刻清零（R56 返修补齐，与空闲相分支对齐）/ clear the instant of the maximum slope, aligned with the idle branch
        _bCross28 := FALSE; // 穿越标志清零 / clear the crossing flag
        _bCross63 := FALSE; // 穿越标志清零 / clear the crossing flag
        _fPvPrev := fPv; // 新基线快照 / take a fresh baseline snapshot
        _fPvBase := fPv; // 新基线过程量 / take a fresh baseline process value
        _eState := E_DL_FopdtState.eRise; // 迁上升相 / migrate to the rise phase
    END_IF

E_DL_FopdtState.eFault: // 故障相：原因锁存，等待复位沿 / fault phase, the cause is latched until the reset edge
    _bValid := FALSE; // 故障拍参数不可交付，数值保持上拍 / parameters are not deliverable and the values hold the last scan

ELSE // 非法相位兜底（R128）/ illegal phase fallback
    _eCause := E_DL_FopdtCause.ePhaseBad; // 成因记非法相位 / record the illegal phase cause
    _bFault := TRUE; // 置故障锁存 / raise the fault latch
    _bValid := FALSE; // 参数不可交付 / parameters not deliverable
    _eState := E_DL_FopdtState.eFault; // 迁故障相 / migrate to the fault phase
END_CASE

// 段 6｜超时判据：仅上升相内判，IN 已带相位闸（R212）/ segment 6, timeout verdict inside the rise phase only, IN already carries the phase gate
IF (_eState = E_DL_FopdtState.eRise) AND tonTimeout.Q AND (NOT _bFault) THEN // 超时且未锁存 / timed out and not yet latched
    _eCause := E_DL_FopdtCause.eNoSettle; // 成因记超时未稳定 / record the timeout without settle cause
    _bFault := TRUE; // 置故障锁存 / raise the fault latch
    _bValid := FALSE; // 参数不可交付 / parameters not deliverable
    _eState := E_DL_FopdtState.eFault; // 迁故障相 / migrate to the fault phase
END_IF

// 段 7｜统一出口：相位映射、单拍脉冲映射、故障锁存与有效位同源 / segment 7, unified outlet for phase mapping, single-shot pulse and matched fault outlets
eState := _eState; // 相位出口单点映射 / single-point phase outlet mapping
eCause := _eCause; // 成因出口单点映射（锁存量）/ single-point cause outlet mapping of the latched value
bError := _bFault; // 故障标志与锁存位同源赋值 / the fault flag shares the latch source
bIdentDone := _bIdentInt; // 完成脉冲映射本拍值 / map the done bit for this scan
_bIdentInt := FALSE; // 映射后立即撤销，保证单拍宽度（R187 两段式）/ revoke right after mapping to keep a single-scan width
bValid := _bValid AND (NOT _bFault); // 有效出口受故障锁存否决（挂状态量，非单拍标志）/ the valid outlet is vetoed by the fault latch, a state quantity
fGainK := _fGainK; // 增益出口 / gain outlet
fTauS := _fTauS; // 时间常数出口 / time constant outlet
fDeadS := _fDeadS; // 纯延迟出口 / dead time outlet
fDeltaPv := _fDeltaPvOut; // 总变化量出口 / total change outlet
fPvBase := _fPvBaseOut; // 基线出口 / baseline outlet
fPvFinal := _fPvFinalOut; // 稳定点出口 / settled value outlet
fTauTwoPointS := _fTauTwoOut; // 两点法时间常数出口 / two-point time constant outlet
fDeadTwoPointS := _fDeadTwoOut; // 两点法纯延迟出口 / two-point dead time outlet
fTauTangentS := _fTauTanOut; // 切线法时间常数出口 / tangent time constant outlet
fDeadTangentS := _fDeadTanOut; // 切线法纯延迟出口 / tangent dead time outlet
END_FUNCTION_BLOCK

(* ---- FB_DL_FrequencyGenerator.st ---- *)
(*
  FB_DL_FrequencyGenerator  —  连续频率发生（方波 + 相位复位 + 占空比组态）/ Continuous frequency generator, square wave
  分类 Category : DL_Algo
  码位 Code     : 16#02_3_86
  段位说明      : 02_3 段占至 85，86 格为 R38 预留解除后的空穴，本件启用 86 格
  版本 Version  : 1.0.0
  来源 Source   : t2-1-lgf-siggen — 信号发生族 R22 已明文分工的「生连续波」侧
  溯源 Origin   : clean-room 实现，相位累加方波发生为公开经典方法，未复制任何源码行
  功能 Function : 1) 连续方波发生：相位累加器 fPhase ∈ [0,1) 每拍推进 fFreqHz * fDt，
                  fPhase < fDuty 为高电平，占空比组态域 [0,1]；
                  2) bPhaseReset 上升沿强制相位归零（多发生器同相启动 / 节拍对齐用）；
                  3) fFreqHz = 0 时输出恒电平：fDuty > 0 恒高、fDuty = 0 恒低（组态级停波）；
                  4) bOutTakenQ 输出本拍电平 + uCycleCnt 周期计数 + fPhaseOut 相位镜像。
  边界 Boundary : ① 与 FB_DL_PulseGenerator 分工：那件是单发/脉宽（发单发），本件是连续波（生连续波）；
                  与 FB_DL_FrequencyMeasure（测）构成「测 ≠ 生」两侧，三件不可互相替代；
                  ② 与 FB_DL_SineGenerator 引脚命名对齐（fFreqHz/fAmplitude/tSampleTime 口径一致）；
                  ③ 无 TON/边沿实例：相位累加器法，任务周期由调用方经 tSampleTime 注入，
                  < T#10MS 钳位（与 FB_DL_RateLimiter 同一口径）；
                  ④ 频率上限钳位 fFreqHzMax：奈奎斯特防御，频率高于任务频率一半时方波失真，
                  越限按上限执行并置信息级码；
                  ⑤ 非有限频率/占空比防御：NaN/Inf 按上次有效值保持，首扫按默认值。
  依赖 Depends  : 仅 Standard.library；与 FB_DL_PulseGenerator / FB_DL_FrequencyMeasure /
                  FB_DL_SineGenerator（均已注册）仅引脚口径对齐，不实例化
  码表 Error codes（本件格 02_3_86，子码步进 +0x100）:
    16#0002_0186 信息级：频率越上限已钳位（奈奎斯特防御，输出按钳后频率执行）
    16#0002_0286 故障级：组态非法（tSampleTime 非正被钳位后仍异常 / 占空比非有限），锁存至 bReset
    16#0002_0386 信息级：相位复位沿生效（fPhase 已归零）

  修订历史 Revision :
    2026-11-19  v1.0.0  R39 首版（批次 1 · 序号 4）
*)

FUNCTION_BLOCK FB_DL_FrequencyGenerator
VAR_INPUT
    bEnable     : BOOL := FALSE;      // 使能，FALSE 时输出恒低并冻结相位 [-] / Enable, FALSE drives output low and freezes phase
    fFreqHz     : REAL := 10.0;       // 目标频率 [Hz]，域 (0, fFreqHzMax]，越限钳位 / Target frequency [Hz], clamped to Nyquist bound
    fDuty       : REAL := 0.5;        // 占空比 [无量纲 0..1]，高电平时间占比 / Duty cycle, high-level fraction
    bPhaseReset : BOOL := FALSE;      // 相位复位，上升沿 fPhase 归零（多路同相启动）/ Phase reset, rising edge zeroes the phase
    bReset      : BOOL := FALSE;      // 故障复位，上升沿清锁存 [-] / Fault reset, rising edge clears latch
    tSampleTime : TIME := T#100MS;    // 任务周期注入 [ms]，< T#10MS 钳位 / Task cycle time injected by caller
END_VAR
VAR_OUTPUT
    bOut        : BOOL;               // 方波输出，TRUE = 高电平相 [-] / Square-wave output, TRUE in high phase
    fPhaseOut   : REAL;               // 相位镜像 [无量纲 0..1)，诊断用 / Phase mirror for diagnostics
    uCycleCnt   : UDINT;              // 输出周期完成计数 [次]，相位回绕一次计一次，饱和 / Completed cycle count, saturating
    bError      : BOOL;               // 故障锁存，仅故障级码置位，bReset 清除 [-] / Fault latch, set only by fault-level codes
    uErrorId    : UDINT;              // 事件码，0 = 无事件（故障级锁存回放）/ Event code, fault codes latched
END_VAR
VAR
    rtPhaseReset : R_TRIG;            // 相位复位沿实例，主体首部无条件刷新 / Phase reset edge instance
    rtReset      : R_TRIG;            // 故障复位沿实例，主体首部无条件刷新 / Fault reset edge instance
    _fPhase      : REAL := 0.0;       // 内部相位累加器 [无量纲 0..1) / Internal phase accumulator
    _fFreqEff    : REAL := 10.0;      // 钳位后的生效频率 [Hz] / Clamped effective frequency
    _fDutyEff    : REAL := 0.5;       // 钳位后的生效占空比 [无量纲] / Clamped effective duty
    _fDt         : REAL := 0.1;       // 生效任务周期 [s] / Effective cycle time in seconds
    _fFreqLast   : REAL := 10.0;      // 上次有效频率保持载体 [Hz]（非有限防御）/ Last valid frequency hold carrier
    _fDutyLast   : REAL := 0.5;       // 上次有效占空比保持载体 [无量纲] / Last valid duty hold carrier
    _bFault      : BOOL;              // 故障锁存位 / Latched fault bit
    _uFault      : UDINT;             // 故障码锁存寄存 / Latched fault code register
    _uInfo       : UDINT;             // 本拍信息码，每拍重算 / Transient info code this cycle
    _bCfgBad     : BOOL;              // 组态非法聚合 / Configuration invalid aggregate
END_VAR
VAR CONSTANT
    DL_FG_DT_MIN     : TIME := T#10MS;      // 任务周期下限钳位 [ms] / Cycle time lower clamp
    DL_FG_FREQ_MAX   : REAL := 50.0;        // 频率组态上限（奈奎斯特防御，按 100ms 任务口径）[Hz] / Frequency configuration bound for Nyquist defense
    DL_FG_INF_CAP    : REAL := 1.0E30;      // 非有限值筛查幅值上限 / Non-finite magnitude screening cap
    DL_FG_CNT_MAX    : UDINT := 16#FFFF_FFFE;  // 周期计数饱和上限 [次] / Cycle count saturation bound
END_VAR

(* —— 段 0：边沿实例无条件周期刷新（R7 红线：严禁置于 IF/CASE 分支内） —— *)
rtPhaseReset(CLK := bPhaseReset);       // 相位复位沿刷新，每拍必调
rtReset(CLK := bReset);                 // 故障复位沿刷新，每拍必调

(* —— 段 1：单拍量预清零（锁存量 _uFault/_bFault 不入清单，R187①） —— *)
_uInfo := 16#0000_0000;                 // 信息码每拍重算
_bCfgBad := FALSE;                      // 组态非法聚合预清零

(* —— 段 2：非有限防御（NaN/Inf 保持上次有效值，首扫用默认） —— *)
IF (fFreqHz <> fFreqHz) OR (ABS(fFreqHz) > DL_FG_INF_CAP) OR ((fFreqHz - fFreqHz) <> 0.0) THEN
    _fFreqEff := _fFreqLast;            // 频率非有限：保持上次有效
    _bCfgBad := TRUE;
ELSE
    _fFreqLast := fFreqHz;              // 有效值入保持载体
    IF fFreqHz < 0.0 THEN
        _fFreqEff := 0.0;               // 负频率钳零（组态级停波）
    ELSIF fFreqHz > DL_FG_FREQ_MAX THEN
        _fFreqEff := DL_FG_FREQ_MAX;    // 越上限钳位（奈奎斯特防御）
        _uInfo := 16#0002_0186;         // 信息级：频率已钳位
    ELSE
        _fFreqEff := fFreqHz;           // 域内直通
    END_IF
END_IF
IF (fDuty <> fDuty) OR (ABS(fDuty) > DL_FG_INF_CAP) OR ((fDuty - fDuty) <> 0.0) THEN
    _fDutyEff := _fDutyLast;            // 占空比非有限：保持上次有效
    _bCfgBad := TRUE;
ELSE
    _fDutyLast := fDuty;
    _fDutyEff := MAX(0.0, MIN(1.0, fDuty));   // 占空比钳到 [0,1]（越界静默钳位，物理量语义）
END_IF

(* —— 段 3：任务周期换算（与 FB_DL_RateLimiter 同口径：< T#10MS 钳位） —— *)
IF tSampleTime < DL_FG_DT_MIN THEN
    _fDt := 0.01;                       // 非法周期钳位 0.01 s
ELSE
    _fDt := TIME_TO_REAL(tSampleTime) / 1000.0;   // TIME 换算秒（显式标准转换）
END_IF

(* —— 段 4：故障锁存与复位沿 —— *)
IF _bCfgBad THEN
    IF NOT _bFault THEN
        _uFault := 16#0002_0286;        // 故障级：组态非法（占空比/频率非有限），仅首次进入时写入
        _bFault := TRUE;
    END_IF
END_IF
IF rtReset.Q THEN
    _bFault := FALSE;                   // 清故障锁存位（唯一解除路径：bReset 上升沿）
    _uFault := 16#0000_0000;
END_IF

(* —— 段 5：相位复位沿（先于推进处理，保证复位拍相位即零） —— *)
IF rtPhaseReset.Q THEN
    _fPhase := 0.0;                     // 相位归零（多路同相启动）
    IF NOT _bFault THEN
        _uInfo := 16#0002_0386;         // 信息级：相位复位生效
    END_IF
END_IF

(* —— 段 6：相位推进与方波生成（失能冻结；故障相保持冻结） —— *)
IF bEnable AND (NOT _bFault) THEN
    _fPhase := _fPhase + _fFreqEff * _fDt;      // 相位推进 = 频率 × 周期
    IF _fPhase >= 1.0 THEN
        _fPhase := _fPhase - 1.0;               // 回绕进位（频率 < 采样率一半时每拍至多进一位）
        uCycleCnt := uCycleCnt + 1;             // 周期完成计数
        IF uCycleCnt >= DL_FG_CNT_MAX THEN
            uCycleCnt := DL_FG_CNT_MAX;         // 计数饱和防回绕
        END_IF
        IF _fPhase >= 1.0 THEN
            _fPhase := 0.0;                     // 极端钳位兜底（频率越限多周回绕）
        END_IF
    END_IF
    bOut := (_fPhase < _fDutyEff);              // 方波判据：相位落在占空比窗内为高电平
END_IF
IF (NOT bEnable) OR _bFault THEN
    bOut := FALSE;                              // 失能/故障：输出恒低（安全侧）
END_IF

(* —— 段 7：出口单点映射（名实同源；锁存码回放，禁同拍抹除） —— *)
fPhaseOut := _fPhase;                           // 相位镜像
IF _bFault THEN
    uErrorId := _uFault;                        // 故障锁存码回放
    bError := TRUE;
ELSE
    uErrorId := _uInfo;                         // 信息码
    bError := FALSE;
END_IF

END_FUNCTION_BLOCK

(* ---- FB_DL_FuzzyTrim2In.st ---- *)
(*==============================================================================
 * 组件名称 (Component)  : FB_DL_FuzzyTrim2In
 * 所属子库 (Sublibrary) : DL_Algo
 * 当前版本 (Version)    : 1.0.0
 * 兼容性   (Platform)   : CODESYS 3.5+ / TwinCAT 3 / 汇川 InoProShop / 施耐德 Machine Expert
 *                         仅依赖 Standard.library（ABS / MAX），零厂商私有库
 * 功能描述 (Function)   : 二输入模糊规则表修调（Mamdani 结构，结构只借、参数自组态）：
 *                         误差 fErr 与误差变化率 fErrRate（均已标幺 -1~1）各做 5 级三角
 *                         隶属度（NB/NS/Z/PS/PB，中心点 -1/-0.5/0/0.5/1，半宽 0.5，
 *                         VAR CONSTANT 可组态）；5×5=25 条规则以 ST_DL_ 常量二维数组落地
 *                         （单点输出集中心，域 [-1,1]）；重心法解模糊：
 *                           fTrim = fGainOut × Σ(w_i×c_i) / Σw_i （w_i = μe×μr）
 *                         适用非线性滞回对象（注塑保压、炉温搭接段）的 PID 外挂修调。
 * 接口     (Interface)  : 输入 fErr 误差（已标幺 -1~1）、fErrRate 误差变化率（已标幺 -1~1）、
 *                         fGainOut 输出增益（>=0）、bReset 复位；输出 fTrim 修调量
 *                         （-fGainOut~+fGainOut）、nRuleHit 命中规则数（诊断）、bNoRule
 *                         无有效规则、bError 组态故障标志。
 * 边界     (Boundary)   : ① **属主边界（写死）：本件只做模糊查表与解模糊，不做标幺换算、
 *                         不接管主回路**；误差/变化率的标幺化由上层标幺件负责。
 *                         ② 输入先钳 [-1,1] 再做隶属度（超域输入不放大）。
 *                         ③ Σw_i 下限闸：Σw_i < 1E-6（全零隶属退化）→ fTrim=0 并置
 *                         bNoRule（防除零，R28）。
 *                         ④ 非有限输入 → 冻结输出（保持上拍 fTrim，不重算）。
 *                         ⑤ 规则表/中心表均为定界常量数组，循环索引为字面常量 0..4，
 *                         天然无越界路径（数组边界红线以静态定界满足）。
 *                         ⑥ 组态闸：fGainOut < 0 → 锁存 bError，输出 0 安全侧，解除沿 =
 *                         bReset 上升沿。
 *                         ⑦ 零全局耦合（无 GVL / 无 VAR_EXTERNAL / 无物理地址）。
 * 分工声明 (Scope)      : 全库无 Fuzzy 族，本件开族；与 PID 族（CascadePid 等）分工：
 *                         模糊修调是非线性补正外挂 ≠ 主调节器。
 * 来源标签 (Source Tag) : T2-5 ◐（Mamdani 结构与重心法只借公开定义，5×5 规则表为本件
 *                         自组态参数域，零文本复制）
 * 码表     (Codes)      : 本件不占用任何全局数字码位。出口为 LREAL 修调量 + BOOL/UDINT 组；
 *                         数字码位待主控收口阶段统一派号。
 * 红线自检 (Redline)    : R1 ✓ 零 GVL/VAR_EXTERNAL ｜ R2 ✓ 零 %I/%Q/%M ｜ R3 ✓ 纯 IEC 61131-3
 *                         R4 ✓ Σw 下限闸 + 输入钳位 + 非有限冻结 ｜ R5 ✓ 声明逐行同行双语注释
 *                         R6 N/A（查表无状态机） ｜ R7 ✓ 一 R_TRIG 段 0 无条件刷新
 * 修订历史 (Revision)   : 2026-11-20  v1.0.0  R48 首版（批次 2 · 序号 8）
 *                         验收向量：e=-1,r=-1 → fTrim=-fGainOut；e=0,r=0 → 0；
 *                         中间值重心插值连续；fGainOut<0 → bError 锁存。
 *==============================================================================*)

TYPE E_DL_FzyTerm :
(
    eNB := 0,    // 负大隶属级 / Negative-big term
    eNS := 1,    // 负小隶属级 / Negative-small term
    eZ  := 2,    // 零隶属级 / Zero term
    ePS := 3,    // 正小隶属级 / Positive-small term
    ePB := 4     // 正大隶属级 / Positive-big term
);
END_TYPE

FUNCTION_BLOCK FB_DL_FuzzyTrim2In
VAR_INPUT
    fErr     : LREAL := 0.0;    // 误差输入（已标幺，域按 [-1,1] 使用，超域先钳） [-] / Error input, normalized
    fErrRate : LREAL := 0.0;    // 误差变化率输入（已标幺） [-] / Error-rate input, normalized
    fGainOut : LREAL := 10.0;   // 修调输出增益（域 >= 0） [工程单位] / Output gain
    bReset   : BOOL := FALSE;   // 复位，上升沿清组态故障锁存 [-] / Reset, rising edge clears config fault
END_VAR
VAR_OUTPUT
    fTrim    : LREAL;           // 模糊修调输出，域 [-fGainOut, +fGainOut] [工程单位] / Fuzzy trim output
    nRuleHit : UDINT;           // 命中规则数（w_i > 0 的规则条数，诊断用） [条] / Rule-hit count for diagnostics
    bNoRule  : BOOL;            // 无有效规则（Σw 过小，输出 0） [-] / No effective rule flag
    bError   : BOOL;            // 组态故障标志（锁存） [-] / Configuration fault flag, latched
END_VAR
VAR
    _fErrC   : LREAL;           // 当拍钳位后误差 [-] / Clamped error this scan
    _fRatC   : LREAL;           // 当拍钳位后误差变化率 [-] / Clamped error rate this scan
    _aMuE    : ARRAY[0..4] OF LREAL;   // 误差五级隶属度 [-] / Error membership grades
    _aMuR    : ARRAY[0..4] OF LREAL;   // 变化率五级隶属度 [-] / Rate membership grades
    _fSumW   : LREAL;           // Σw 累加中间量 [-] / Weight sum accumulator
    _fSumWC  : LREAL;           // Σ(w×c) 累加中间量 [-] / Weighted-center accumulator
    _nHit    : UDINT;           // 命中规则内部量 [条] / Rule-hit internal
    _fTrim   : LREAL := 0.0;    // 修调锁存镜像（冻结源） / Trim latch mirror, freeze source
    _bErrLatch : BOOL;          // 组态故障锁存位（解除沿 = bReset 上升沿） / Latched config fault, cleared by reset edge
    rtReset  : R_TRIG;          // 复位沿实例，段 0 无条件调用 / Reset edge instance
    _bNonFin : BOOL;            // 输入非有限当拍量 [-] / Non-finite input this scan
    i        : DINT;            // 规则表行索引（误差级） / Rule table row index
    j        : DINT;            // 规则表列索引（变化率级） / Rule table column index
    _fW      : LREAL;           // 单规则权重中间量 [-] / Single rule weight
END_VAR
VAR CONSTANT
    DL_FZY_HALF  : LREAL := 0.5;      // 三角隶属半宽（中心间隔相同） [-] / Triangle membership half-width
    DL_FZY_WMIN  : LREAL := 1.0E-6;   // Σw 下限闸（防除零） [-] / Weight-sum floor
    DL_FZY_ONE   : LREAL := 1.0;      // 单位常量（钳位上限） [-] / Unit constant
    DL_FZY_CEN   : ARRAY[0..4] OF LREAL := [-1.0, -0.5, 0.0, 0.5, 1.0];   // 五级隶属中心点（NB/NS/Z/PS/PB），组态参数域 [-] / Five membership centers
    DL_FZY_RULE  : ARRAY[0..4, 0..4] OF LREAL := [   // 5×5 规则表：行=误差级、列=变化率级 [-] / 5x5 rule table of singleton centers
        -1.0, -1.0, -0.5, -0.5,  0.0,
        -1.0, -0.5, -0.5,  0.0,  0.5,
        -0.5, -0.5,  0.0,  0.5,  0.5,
        -0.5,  0.0,  0.5,  0.5,  1.0,
         0.0,  0.5,  0.5,  1.0,  1.0];
                                      // 5×5 规则表：行=误差级、列=变化率级，值为单点输出集中心，对称反对角设计 [-] / 5x5 rule table of singleton centers
END_VAR

(* —— 段 0：非有限判 + 组态闸 + 输入钳位 + 沿刷新 —— *)
_bNonFin := (fErr <> fErr) OR ((fErr - fErr) <> 0.0)
         OR (fErrRate <> fErrRate) OR ((fErrRate - fErrRate) <> 0.0);   // 输入非有限（R245） / Non-finite input tests
IF fGainOut < 0.0 THEN
    _bErrLatch := TRUE;                                   // 增益负值组态闸：锁存（R188 解除沿 = bReset 上升沿） / Negative gain gate: latch
END_IF
rtReset(CLK := bReset);                                   // 复位沿，每拍必调 / Reset edge, every scan

(* —— 段 1：复位沿 —— *)
IF rtReset.Q THEN
    _bErrLatch := FALSE;                                  // 清组态故障锁存 / Clear config fault latch
END_IF

(* —— 段 2：隶属度与解模糊（非有限冻结；故障期安全侧） —— *)
nRuleHit := 0;                                            // 命中数出口预清 / Hit count preset
bNoRule  := FALSE;                                        // 无规则标志预清 / No-rule flag preset
IF _bErrLatch THEN
    _fTrim := 0.0;                                        // 故障安全侧：修调归零 / Fault safe side: zero trim
ELSIF _bNonFin THEN
    (* 非有限输入：冻结上拍 _fTrim 不重算（头注释④） *)
    ;                                                     // 冻结分支保持 / Freeze branch holds
ELSE
    IF fErr > DL_FZY_ONE THEN
        _fErrC := DL_FZY_ONE;                             // 误差上钳 [-1,1] / Clamp error high
    ELSIF fErr < -DL_FZY_ONE THEN
        _fErrC := -DL_FZY_ONE;                            // 误差下钳 / Clamp error low
    ELSE
        _fErrC := fErr;                                   // 域内直通 / In-domain pass
    END_IF
    IF fErrRate > DL_FZY_ONE THEN
        _fRatC := DL_FZY_ONE;                             // 变化率上钳 / Clamp rate high
    ELSIF fErrRate < -DL_FZY_ONE THEN
        _fRatC := -DL_FZY_ONE;                            // 变化率下钳 / Clamp rate low
    ELSE
        _fRatC := fErrRate;                               // 域内直通 / In-domain pass
    END_IF
    FOR i := 0 TO 4 DO
        IF (_fErrC - DL_FZY_CEN[i]) < 0.0 THEN
            _aMuE[i] := DL_FZY_HALF + (_fErrC - DL_FZY_CEN[i]);   // 左斜坡隶属（三角左半）/ Left ramp membership
        ELSE
            _aMuE[i] := DL_FZY_HALF - (_fErrC - DL_FZY_CEN[i]);   // 右斜坡隶属（三角右半）/ Right ramp membership
        END_IF
        IF _aMuE[i] < 0.0 THEN
            _aMuE[i] := 0.0;                              // 负隶属截零 / Clamp membership to zero
        END_IF
        IF (_fRatC - DL_FZY_CEN[i]) < 0.0 THEN
            _aMuR[i] := DL_FZY_HALF + (_fRatC - DL_FZY_CEN[i]);   // 变化率左斜坡 / Rate left ramp
        ELSE
            _aMuR[i] := DL_FZY_HALF - (_fRatC - DL_FZY_CEN[i]);   // 变化率右斜坡 / Rate right ramp
        END_IF
        IF _aMuR[i] < 0.0 THEN
            _aMuR[i] := 0.0;                              // 负隶属截零 / Clamp membership to zero
        END_IF
    END_FOR
    _fSumW  := 0.0;                                       // Σw 清零 / Clear weight sum
    _fSumWC := 0.0;                                       // Σ(w×c) 清零 / Clear weighted center
    _nHit   := 0;                                         // 命中数清零 / Clear hit count
    FOR i := 0 TO 4 DO
        FOR j := 0 TO 4 DO
            _fW := _aMuE[i] * _aMuR[j];                   // 单规则权重 = μe×μr / Single rule weight
            IF _fW > 0.0 THEN
                _fSumW  := _fSumW + _fW;                  // 累加权重 / Accumulate weight
                _fSumWC := _fSumWC + _fW * DL_FZY_RULE[i][j];   // 累加权重×中心 / Accumulate weight times center
                _nHit := _nHit + 1;                       // 命中规则计数 / Count hit rule
            END_IF
        END_FOR
    END_FOR
    IF _fSumW < DL_FZY_WMIN THEN
        _fTrim := 0.0;                                    // Σw 下限闸：全零隶属退化输出 0（R28 防除零） / Weight-sum floor: zero output
        bNoRule := TRUE;                                  // 置无有效规则标志 / Raise no-rule flag
        _nHit := 0;                                       // 无有效规则命中数归零 / Zero hit count
    ELSE
        _fTrim := fGainOut * _fSumWC / _fSumW;            // 重心法解模糊（分母已过闸） / Centre-of-gravity defuzzification
    END_IF
END_IF

(* —— 段 3：出口单点映射（名实双出口同源，R191） —— *)
fTrim    := _fTrim;                                       // 修调出口 / Trim outlet
nRuleHit := _nHit;                                        // 命中数出口 / Hit count outlet
bError   := _bErrLatch;                                   // 故障标志出口 / Error flag outlet

END_FUNCTION_BLOCK
